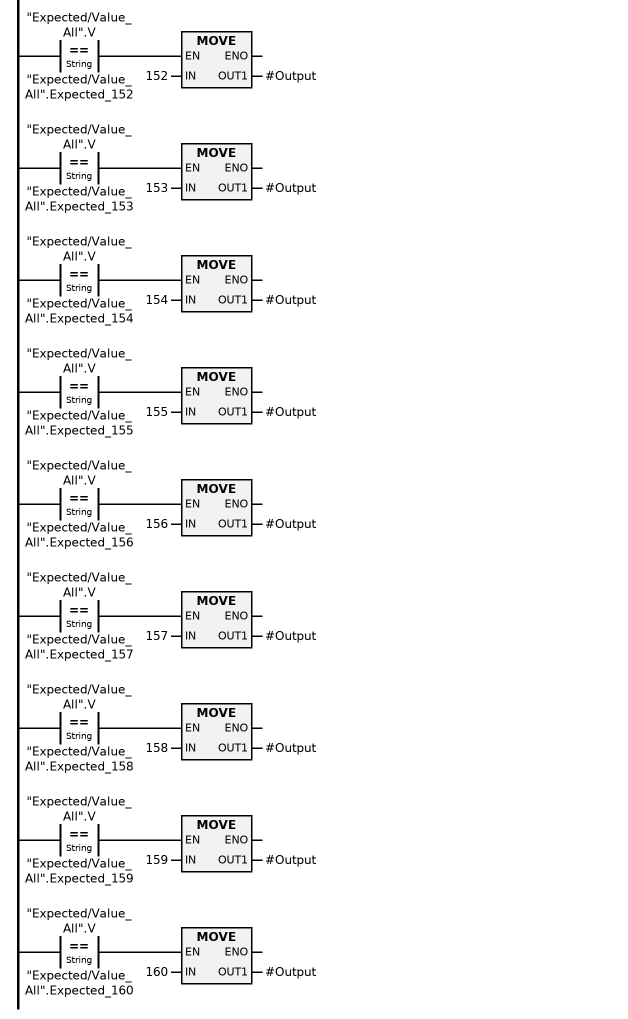
   RUNG wire#powerrail
      { S7_Templates := "SrcType := String" } EQ_Contact(in1 := "Expected/Value_All".V, in2 := "Expected/Value_All".Expected_141)
      Move(in := 141, out1 => #Output)
   END_RUNG
   RUNG wire#powerrail
      { S7_Templates := "SrcType := String" } EQ_Contact(in1 := "Expected/Value_All".V, in2 := "Expected/Value_All".Expected_142)
      Move(in := 142, out1 => #Output)
   END_RUNG
   RUNG wire#powerrail
      { S7_Templates := "SrcType := String" } EQ_Contact(in1 := "Expected/Value_All".V, in2 := "Expected/Value_All".Expected_143)
      Move(in := 143, out1 => #Output)
   END_RUNG
   RUNG wire#powerrail
      { S7_Templates := "SrcType := String" } EQ_Contact(in1 := "Expected/Value_All".V, in2 := "Expected/Value_All".Expected_144)
      Move(in := 144, out1 => #Output)
   END_RUNG
   RUNG wire#powerrail
      { S7_Templates := "SrcType := String" } EQ_Contact(in1 := "Expected/Value_All".V, in2 := "Expected/Value_All".Expected_145)
      Move(in := 145, out1 => #Output)
   END_RUNG
   RUNG wire#powerrail
      { S7_Templates := "SrcType := String" } EQ_Contact(in1 := "Expected/Value_All".V, in2 := "Expected/Value_All".Expected_146)
      Move(in := 146, out1 => #Output)
   END_RUNG
   RUNG wire#powerrail
      { S7_Templates := "SrcType := String" } EQ_Contact(in1 := "Expected/Value_All".V, in2 := "Expected/Value_All".Expected_147)
      Move(in := 147, out1 => #Output)
   END_RUNG
   RUNG wire#powerrail
      { S7_Templates := "SrcType := String" } EQ_Contact(in1 := "Expected/Value_All".V, in2 := "Expected/Value_All".Expected_148)
      Move(in := 148, out1 => #Output)
   END_RUNG
   RUNG wire#powerrail
      { S7_Templates := "SrcType := String" } EQ_Contact(in1 := "Expected/Value_All".V, in2 := "Expected/Value_All".Expected_149)
      Move(in := 149, out1 => #Output)
   END_RUNG
   RUNG wire#powerrail
      { S7_Templates := "SrcType := String" } EQ_Contact(in1 := "Expected/Value_All".V, in2 := "Expected/Value_All".Expected_150)
      Move(in := 150, out1 => #Output)
   END_RUNG
   RUNG wire#powerrail
      { S7_Templates := "SrcType := String" } EQ_Contact(in1 := "Expected/Value_All".V, in2 := "Expected/Value_All".Expected_151)
      Move(in := 151, out1 => #Output)
   END_RUNG
   RUNG wire#powerrail
      { S7_Templates := "SrcType := String" } EQ_Contact(in1 := "Expected/Value_All".V, in2 := "Expected/Value_All".Expected_152)
      Move(in := 152, out1 => #Output)
   END_RUNG
   RUNG wire#powerrail
      { S7_Templates := "SrcType := String" } EQ_Contact(in1 := "Expected/Value_All".V, in2 := "Expected/Value_All".Expected_153)
      Move(in := 153, out1 => #Output)
   END_RUNG
   RUNG wire#powerrail
      { S7_Templates := "SrcType := String" } EQ_Contact(in1 := "Expected/Value_All".V, in2 := "Expected/Value_All".Expected_154)
      Move(in := 154, out1 => #Output)
   END_RUNG
   RUNG wire#powerrail
      { S7_Templates := "SrcType := String" } EQ_Contact(in1 := "Expected/Value_All".V, in2 := "Expected/Value_All".Expected_155)
      Move(in := 155, out1 => #Output)
   END_RUNG
   RUNG wire#powerrail
      { S7_Templates := "SrcType := String" } EQ_Contact(in1 := "Expected/Value_All".V, in2 := "Expected/Value_All".Expected_156)
      Move(in := 156, out1 => #Output)
   END_RUNG
   RUNG wire#powerrail
      { S7_Templates := "SrcType := String" } EQ_Contact(in1 := "Expected/Value_All".V, in2 := "Expected/Value_All".Expected_157)
      Move(in := 157, out1 => #Output)
   END_RUNG
   RUNG wire#powerrail
      { S7_Templates := "SrcType := String" } EQ_Contact(in1 := "Expected/Value_All".V, in2 := "Expected/Value_All".Expected_158)
      Move(in := 158, out1 => #Output)
   END_RUNG
   RUNG wire#powerrail
      { S7_Templates := "SrcType := String" } EQ_Contact(in1 := "Expected/Value_All".V, in2 := "Expected/Value_All".Expected_159)
      Move(in := 159, out1 => #Output)
   END_RUNG
   RUNG wire#powerrail
      { S7_Templates := "SrcType := String" } EQ_Contact(in1 := "Expected/Value_All".V, in2 := "Expected/Value_All".Expected_160)
      Move(in := 160, out1 => #Output)
   END_RUNG
   // the same network as SCL:
   IF "Expected/Value_All".V = "Expected/Value_All".Expected_141 THEN #Output := 141; END_IF;
   IF "Expected/Value_All".V = "Expected/Value_All".Expected_142 THEN #Output := 142; END_IF;
   IF "Expected/Value_All".V = "Expected/Value_All".Expected_143 THEN #Output := 143; END_IF;
   IF "Expected/Value_All".V = "Expected/Value_All".Expected_144 THEN #Output := 144; END_IF;
   IF "Expected/Value_All".V = "Expected/Value_All".Expected_145 THEN #Output := 145; END_IF;
   IF "Expected/Value_All".V = "Expected/Value_All".Expected_146 THEN #Output := 146; END_IF;
   IF "Expected/Value_All".V = "Expected/Value_All".Expected_147 THEN #Output := 147; END_IF;
   IF "Expected/Value_All".V = "Expected/Value_All".Expected_148 THEN #Output := 148; END_IF;
   IF "Expected/Value_All".V = "Expected/Value_All".Expected_149 THEN #Output := 149; END_IF;
   IF "Expected/Value_All".V = "Expected/Value_All".Expected_150 THEN #Output := 150; END_IF;
   IF "Expected/Value_All".V = "Expected/Value_All".Expected_151 THEN #Output := 151; END_IF;
   IF "Expected/Value_All".V = "Expected/Value_All".Expected_152 THEN #Output := 152; END_IF;
   IF "Expected/Value_All".V = "Expected/Value_All".Expected_153 THEN #Output := 153; END_IF;
   IF "Expected/Value_All".V = "Expected/Value_All".Expected_154 THEN #Output := 154; END_IF;
   IF "Expected/Value_All".V = "Expected/Value_All".Expected_155 THEN #Output := 155; END_IF;
   IF "Expected/Value_All".V = "Expected/Value_All".Expected_156 THEN #Output := 156; END_IF;
   IF "Expected/Value_All".V = "Expected/Value_All".Expected_157 THEN #Output := 157; END_IF;
   IF "Expected/Value_All".V = "Expected/Value_All".Expected_158 THEN #Output := 158; END_IF;
   IF "Expected/Value_All".V = "Expected/Value_All".Expected_159 THEN #Output := 159; END_IF;
   IF "Expected/Value_All".V = "Expected/Value_All".Expected_160 THEN #Output := 160; END_IF;
END_REGION

REGION Network 9
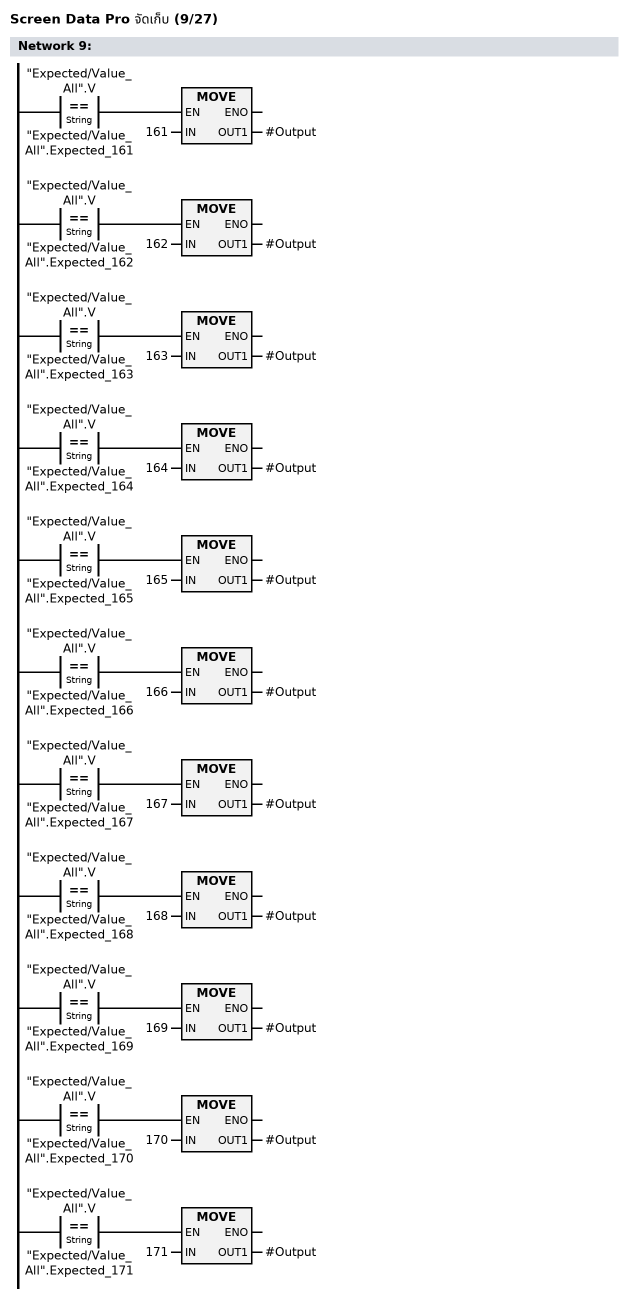
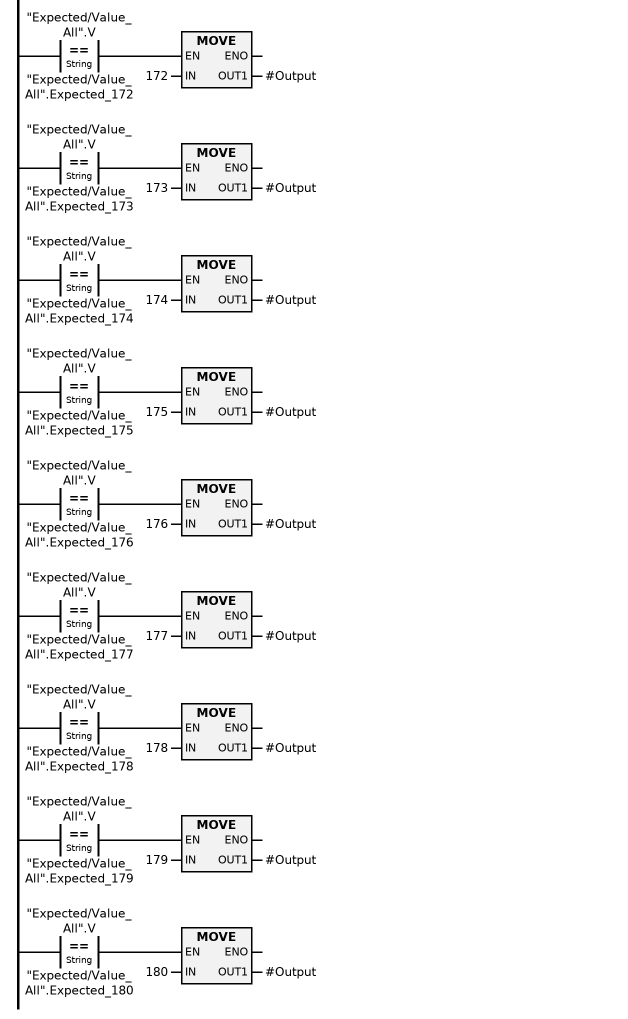
   RUNG wire#powerrail
      { S7_Templates := "SrcType := String" } EQ_Contact(in1 := "Expected/Value_All".V, in2 := "Expected/Value_All".Expected_161)
      Move(in := 161, out1 => #Output)
   END_RUNG
   RUNG wire#powerrail
      { S7_Templates := "SrcType := String" } EQ_Contact(in1 := "Expected/Value_All".V, in2 := "Expected/Value_All".Expected_162)
      Move(in := 162, out1 => #Output)
   END_RUNG
   RUNG wire#powerrail
      { S7_Templates := "SrcType := String" } EQ_Contact(in1 := "Expected/Value_All".V, in2 := "Expected/Value_All".Expected_163)
      Move(in := 163, out1 => #Output)
   END_RUNG
   RUNG wire#powerrail
      { S7_Templates := "SrcType := String" } EQ_Contact(in1 := "Expected/Value_All".V, in2 := "Expected/Value_All".Expected_164)
      Move(in := 164, out1 => #Output)
   END_RUNG
   RUNG wire#powerrail
      { S7_Templates := "SrcType := String" } EQ_Contact(in1 := "Expected/Value_All".V, in2 := "Expected/Value_All".Expected_165)
      Move(in := 165, out1 => #Output)
   END_RUNG
   RUNG wire#powerrail
      { S7_Templates := "SrcType := String" } EQ_Contact(in1 := "Expected/Value_All".V, in2 := "Expected/Value_All".Expected_166)
      Move(in := 166, out1 => #Output)
   END_RUNG
   RUNG wire#powerrail
      { S7_Templates := "SrcType := String" } EQ_Contact(in1 := "Expected/Value_All".V, in2 := "Expected/Value_All".Expected_167)
      Move(in := 167, out1 => #Output)
   END_RUNG
   RUNG wire#powerrail
      { S7_Templates := "SrcType := String" } EQ_Contact(in1 := "Expected/Value_All".V, in2 := "Expected/Value_All".Expected_168)
      Move(in := 168, out1 => #Output)
   END_RUNG
   RUNG wire#powerrail
      { S7_Templates := "SrcType := String" } EQ_Contact(in1 := "Expected/Value_All".V, in2 := "Expected/Value_All".Expected_169)
      Move(in := 169, out1 => #Output)
   END_RUNG
   RUNG wire#powerrail
      { S7_Templates := "SrcType := String" } EQ_Contact(in1 := "Expected/Value_All".V, in2 := "Expected/Value_All".Expected_170)
      Move(in := 170, out1 => #Output)
   END_RUNG
   RUNG wire#powerrail
      { S7_Templates := "SrcType := String" } EQ_Contact(in1 := "Expected/Value_All".V, in2 := "Expected/Value_All".Expected_171)
      Move(in := 171, out1 => #Output)
   END_RUNG
   RUNG wire#powerrail
      { S7_Templates := "SrcType := String" } EQ_Contact(in1 := "Expected/Value_All".V, in2 := "Expected/Value_All".Expected_172)
      Move(in := 172, out1 => #Output)
   END_RUNG
   RUNG wire#powerrail
      { S7_Templates := "SrcType := String" } EQ_Contact(in1 := "Expected/Value_All".V, in2 := "Expected/Value_All".Expected_173)
      Move(in := 173, out1 => #Output)
   END_RUNG
   RUNG wire#powerrail
      { S7_Templates := "SrcType := String" } EQ_Contact(in1 := "Expected/Value_All".V, in2 := "Expected/Value_All".Expected_174)
      Move(in := 174, out1 => #Output)
   END_RUNG
   RUNG wire#powerrail
      { S7_Templates := "SrcType := String" } EQ_Contact(in1 := "Expected/Value_All".V, in2 := "Expected/Value_All".Expected_175)
      Move(in := 175, out1 => #Output)
   END_RUNG
   RUNG wire#powerrail
      { S7_Templates := "SrcType := String" } EQ_Contact(in1 := "Expected/Value_All".V, in2 := "Expected/Value_All".Expected_176)
      Move(in := 176, out1 => #Output)
   END_RUNG
   RUNG wire#powerrail
      { S7_Templates := "SrcType := String" } EQ_Contact(in1 := "Expected/Value_All".V, in2 := "Expected/Value_All".Expected_177)
      Move(in := 177, out1 => #Output)
   END_RUNG
   RUNG wire#powerrail
      { S7_Templates := "SrcType := String" } EQ_Contact(in1 := "Expected/Value_All".V, in2 := "Expected/Value_All".Expected_178)
      Move(in := 178, out1 => #Output)
   END_RUNG
   RUNG wire#powerrail
      { S7_Templates := "SrcType := String" } EQ_Contact(in1 := "Expected/Value_All".V, in2 := "Expected/Value_All".Expected_179)
      Move(in := 179, out1 => #Output)
   END_RUNG
   RUNG wire#powerrail
      { S7_Templates := "SrcType := String" } EQ_Contact(in1 := "Expected/Value_All".V, in2 := "Expected/Value_All".Expected_180)
      Move(in := 180, out1 => #Output)
   END_RUNG
   // the same network as SCL:
   IF "Expected/Value_All".V = "Expected/Value_All".Expected_161 THEN #Output := 161; END_IF;
   IF "Expected/Value_All".V = "Expected/Value_All".Expected_162 THEN #Output := 162; END_IF;
   IF "Expected/Value_All".V = "Expected/Value_All".Expected_163 THEN #Output := 163; END_IF;
   IF "Expected/Value_All".V = "Expected/Value_All".Expected_164 THEN #Output := 164; END_IF;
   IF "Expected/Value_All".V = "Expected/Value_All".Expected_165 THEN #Output := 165; END_IF;
   IF "Expected/Value_All".V = "Expected/Value_All".Expected_166 THEN #Output := 166; END_IF;
   IF "Expected/Value_All".V = "Expected/Value_All".Expected_167 THEN #Output := 167; END_IF;
   IF "Expected/Value_All".V = "Expected/Value_All".Expected_168 THEN #Output := 168; END_IF;
   IF "Expected/Value_All".V = "Expected/Value_All".Expected_169 THEN #Output := 169; END_IF;
   IF "Expected/Value_All".V = "Expected/Value_All".Expected_170 THEN #Output := 170; END_IF;
   IF "Expected/Value_All".V = "Expected/Value_All".Expected_171 THEN #Output := 171; END_IF;
   IF "Expected/Value_All".V = "Expected/Value_All".Expected_172 THEN #Output := 172; END_IF;
   IF "Expected/Value_All".V = "Expected/Value_All".Expected_173 THEN #Output := 173; END_IF;
   IF "Expected/Value_All".V = "Expected/Value_All".Expected_174 THEN #Output := 174; END_IF;
   IF "Expected/Value_All".V = "Expected/Value_All".Expected_175 THEN #Output := 175; END_IF;
   IF "Expected/Value_All".V = "Expected/Value_All".Expected_176 THEN #Output := 176; END_IF;
   IF "Expected/Value_All".V = "Expected/Value_All".Expected_177 THEN #Output := 177; END_IF;
   IF "Expected/Value_All".V = "Expected/Value_All".Expected_178 THEN #Output := 178; END_IF;
   IF "Expected/Value_All".V = "Expected/Value_All".Expected_179 THEN #Output := 179; END_IF;
   IF "Expected/Value_All".V = "Expected/Value_All".Expected_180 THEN #Output := 180; END_IF;
END_REGION

REGION Network 10
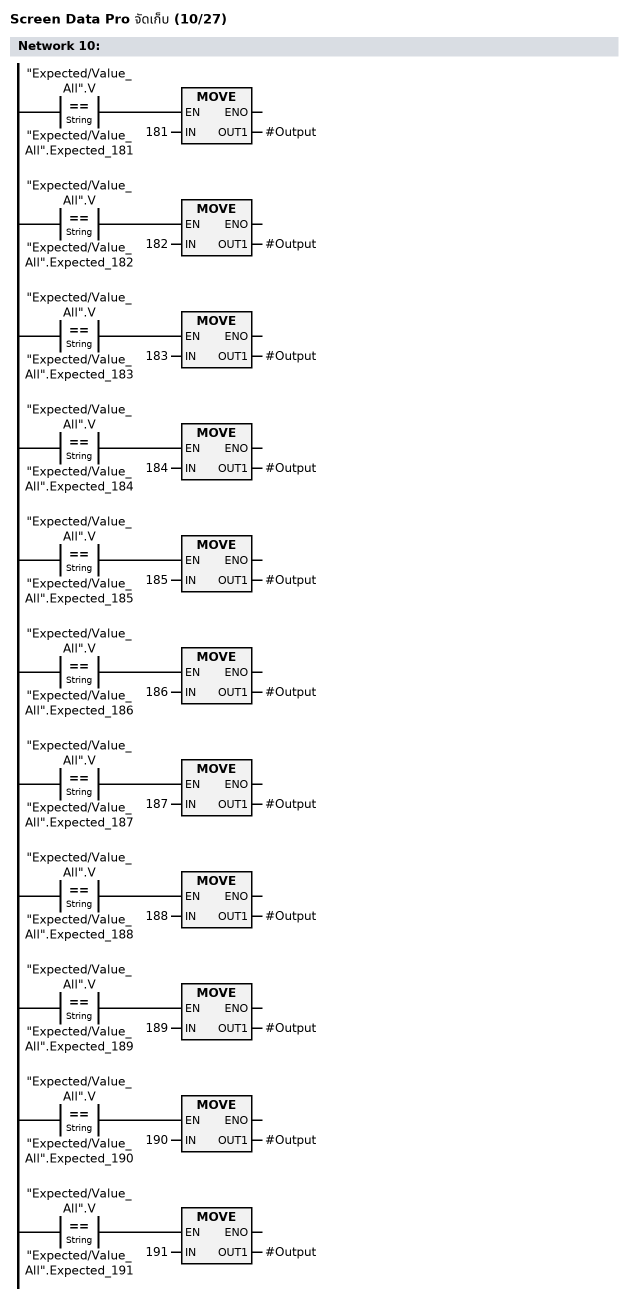
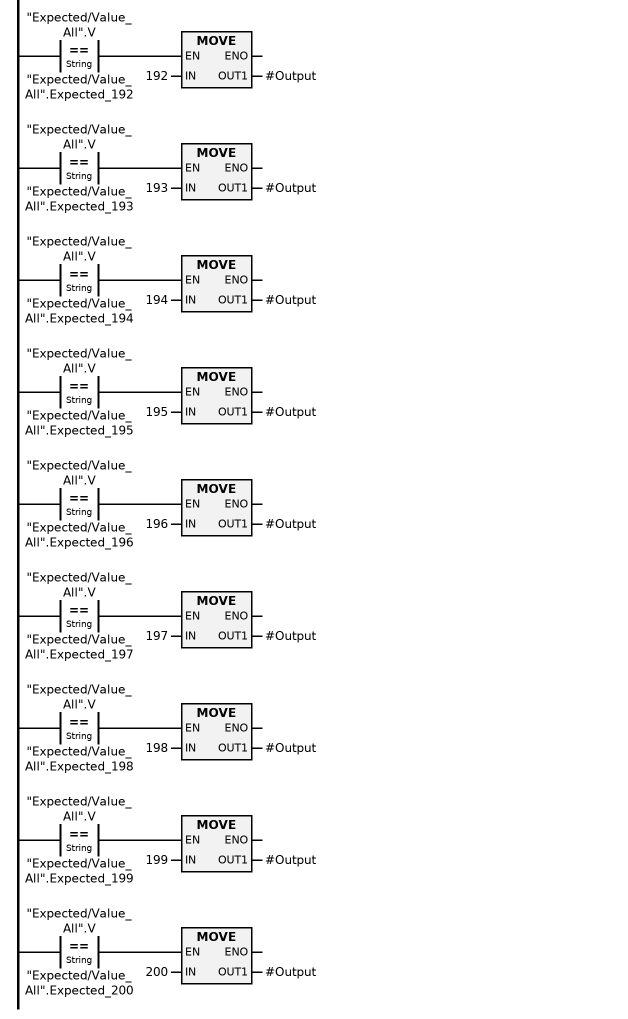
   RUNG wire#powerrail
      { S7_Templates := "SrcType := String" } EQ_Contact(in1 := "Expected/Value_All".V, in2 := "Expected/Value_All".Expected_181)
      Move(in := 181, out1 => #Output)
   END_RUNG
   RUNG wire#powerrail
      { S7_Templates := "SrcType := String" } EQ_Contact(in1 := "Expected/Value_All".V, in2 := "Expected/Value_All".Expected_182)
      Move(in := 182, out1 => #Output)
   END_RUNG
   RUNG wire#powerrail
      { S7_Templates := "SrcType := String" } EQ_Contact(in1 := "Expected/Value_All".V, in2 := "Expected/Value_All".Expected_183)
      Move(in := 183, out1 => #Output)
   END_RUNG
   RUNG wire#powerrail
      { S7_Templates := "SrcType := String" } EQ_Contact(in1 := "Expected/Value_All".V, in2 := "Expected/Value_All".Expected_184)
      Move(in := 184, out1 => #Output)
   END_RUNG
   RUNG wire#powerrail
      { S7_Templates := "SrcType := String" } EQ_Contact(in1 := "Expected/Value_All".V, in2 := "Expected/Value_All".Expected_185)
      Move(in := 185, out1 => #Output)
   END_RUNG
   RUNG wire#powerrail
      { S7_Templates := "SrcType := String" } EQ_Contact(in1 := "Expected/Value_All".V, in2 := "Expected/Value_All".Expected_186)
      Move(in := 186, out1 => #Output)
   END_RUNG
   RUNG wire#powerrail
      { S7_Templates := "SrcType := String" } EQ_Contact(in1 := "Expected/Value_All".V, in2 := "Expected/Value_All".Expected_187)
      Move(in := 187, out1 => #Output)
   END_RUNG
   RUNG wire#powerrail
      { S7_Templates := "SrcType := String" } EQ_Contact(in1 := "Expected/Value_All".V, in2 := "Expected/Value_All".Expected_188)
      Move(in := 188, out1 => #Output)
   END_RUNG
   RUNG wire#powerrail
      { S7_Templates := "SrcType := String" } EQ_Contact(in1 := "Expected/Value_All".V, in2 := "Expected/Value_All".Expected_189)
      Move(in := 189, out1 => #Output)
   END_RUNG
   RUNG wire#powerrail
      { S7_Templates := "SrcType := String" } EQ_Contact(in1 := "Expected/Value_All".V, in2 := "Expected/Value_All".Expected_190)
      Move(in := 190, out1 => #Output)
   END_RUNG
   RUNG wire#powerrail
      { S7_Templates := "SrcType := String" } EQ_Contact(in1 := "Expected/Value_All".V, in2 := "Expected/Value_All".Expected_191)
      Move(in := 191, out1 => #Output)
   END_RUNG
   RUNG wire#powerrail
      { S7_Templates := "SrcType := String" } EQ_Contact(in1 := "Expected/Value_All".V, in2 := "Expected/Value_All".Expected_192)
      Move(in := 192, out1 => #Output)
   END_RUNG
   RUNG wire#powerrail
      { S7_Templates := "SrcType := String" } EQ_Contact(in1 := "Expected/Value_All".V, in2 := "Expected/Value_All".Expected_193)
      Move(in := 193, out1 => #Output)
   END_RUNG
   RUNG wire#powerrail
      { S7_Templates := "SrcType := String" } EQ_Contact(in1 := "Expected/Value_All".V, in2 := "Expected/Value_All".Expected_194)
      Move(in := 194, out1 => #Output)
   END_RUNG
   RUNG wire#powerrail
      { S7_Templates := "SrcType := String" } EQ_Contact(in1 := "Expected/Value_All".V, in2 := "Expected/Value_All".Expected_195)
      Move(in := 195, out1 => #Output)
   END_RUNG
   RUNG wire#powerrail
      { S7_Templates := "SrcType := String" } EQ_Contact(in1 := "Expected/Value_All".V, in2 := "Expected/Value_All".Expected_196)
      Move(in := 196, out1 => #Output)
   END_RUNG
   RUNG wire#powerrail
      { S7_Templates := "SrcType := String" } EQ_Contact(in1 := "Expected/Value_All".V, in2 := "Expected/Value_All".Expected_197)
      Move(in := 197, out1 => #Output)
   END_RUNG
   RUNG wire#powerrail
      { S7_Templates := "SrcType := String" } EQ_Contact(in1 := "Expected/Value_All".V, in2 := "Expected/Value_All".Expected_198)
      Move(in := 198, out1 => #Output)
   END_RUNG
   RUNG wire#powerrail
      { S7_Templates := "SrcType := String" } EQ_Contact(in1 := "Expected/Value_All".V, in2 := "Expected/Value_All".Expected_199)
      Move(in := 199, out1 => #Output)
   END_RUNG
   RUNG wire#powerrail
      { S7_Templates := "SrcType := String" } EQ_Contact(in1 := "Expected/Value_All".V, in2 := "Expected/Value_All".Expected_200)
      Move(in := 200, out1 => #Output)
   END_RUNG
   // the same network as SCL:
   IF "Expected/Value_All".V = "Expected/Value_All".Expected_181 THEN #Output := 181; END_IF;
   IF "Expected/Value_All".V = "Expected/Value_All".Expected_182 THEN #Output := 182; END_IF;
   IF "Expected/Value_All".V = "Expected/Value_All".Expected_183 THEN #Output := 183; END_IF;
   IF "Expected/Value_All".V = "Expected/Value_All".Expected_184 THEN #Output := 184; END_IF;
   IF "Expected/Value_All".V = "Expected/Value_All".Expected_185 THEN #Output := 185; END_IF;
   IF "Expected/Value_All".V = "Expected/Value_All".Expected_186 THEN #Output := 186; END_IF;
   IF "Expected/Value_All".V = "Expected/Value_All".Expected_187 THEN #Output := 187; END_IF;
   IF "Expected/Value_All".V = "Expected/Value_All".Expected_188 THEN #Output := 188; END_IF;
   IF "Expected/Value_All".V = "Expected/Value_All".Expected_189 THEN #Output := 189; END_IF;
   IF "Expected/Value_All".V = "Expected/Value_All".Expected_190 THEN #Output := 190; END_IF;
   IF "Expected/Value_All".V = "Expected/Value_All".Expected_191 THEN #Output := 191; END_IF;
   IF "Expected/Value_All".V = "Expected/Value_All".Expected_192 THEN #Output := 192; END_IF;
   IF "Expected/Value_All".V = "Expected/Value_All".Expected_193 THEN #Output := 193; END_IF;
   IF "Expected/Value_All".V = "Expected/Value_All".Expected_194 THEN #Output := 194; END_IF;
   IF "Expected/Value_All".V = "Expected/Value_All".Expected_195 THEN #Output := 195; END_IF;
   IF "Expected/Value_All".V = "Expected/Value_All".Expected_196 THEN #Output := 196; END_IF;
   IF "Expected/Value_All".V = "Expected/Value_All".Expected_197 THEN #Output := 197; END_IF;
   IF "Expected/Value_All".V = "Expected/Value_All".Expected_198 THEN #Output := 198; END_IF;
   IF "Expected/Value_All".V = "Expected/Value_All".Expected_199 THEN #Output := 199; END_IF;
   IF "Expected/Value_All".V = "Expected/Value_All".Expected_200 THEN #Output := 200; END_IF;
END_REGION

REGION Network 11
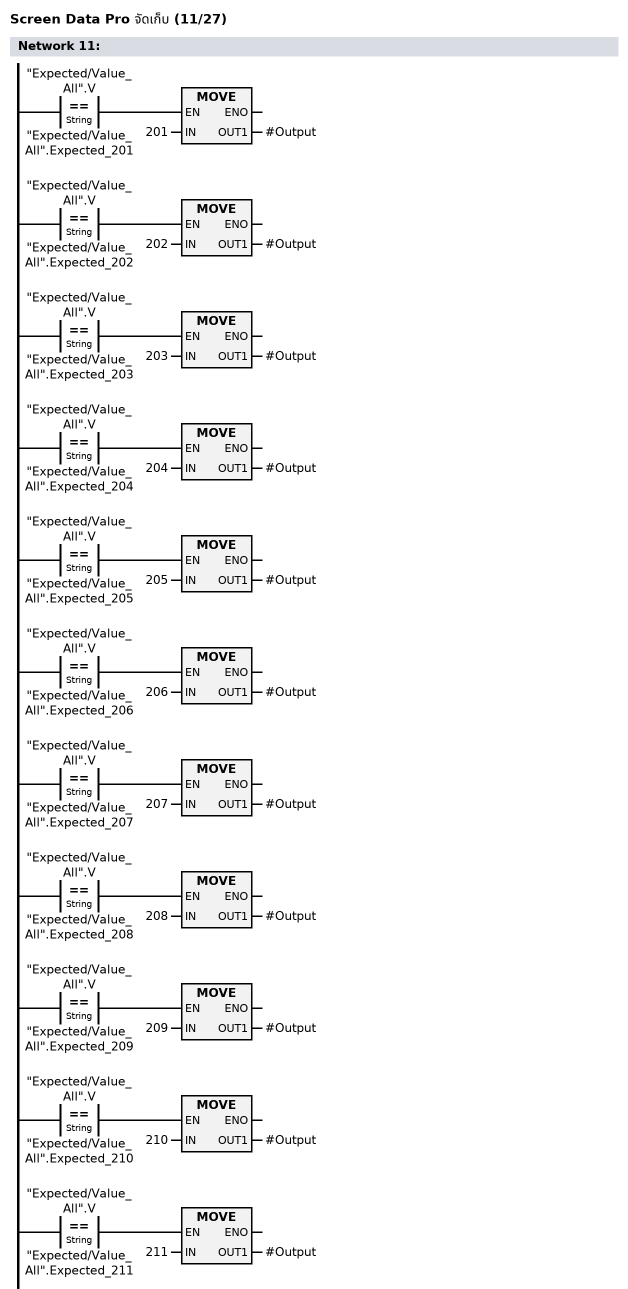
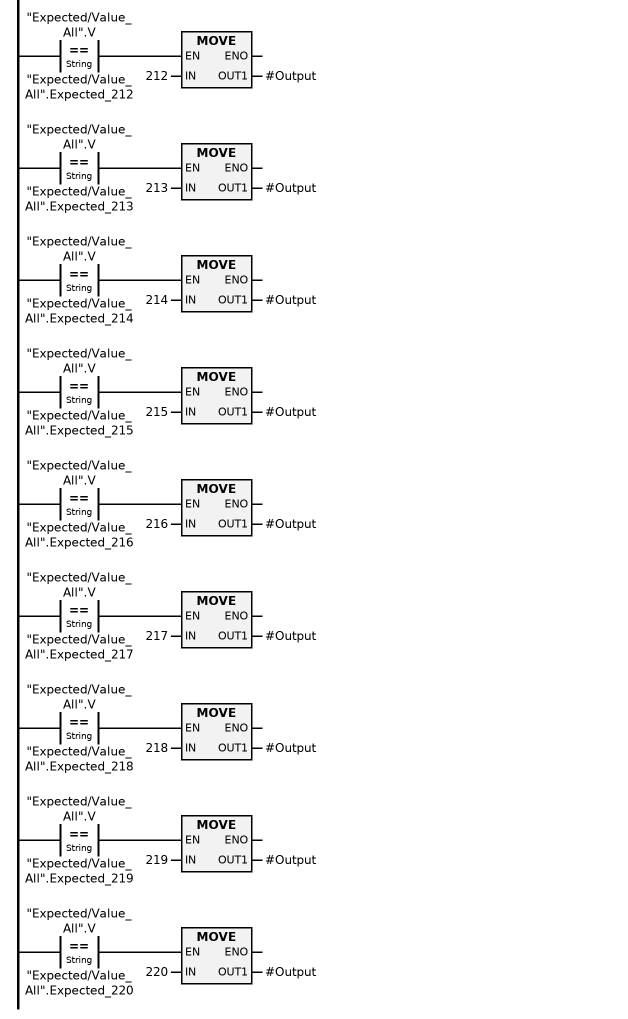
   RUNG wire#powerrail
      { S7_Templates := "SrcType := String" } EQ_Contact(in1 := "Expected/Value_All".V, in2 := "Expected/Value_All".Expected_201)
      Move(in := 201, out1 => #Output)
   END_RUNG
   RUNG wire#powerrail
      { S7_Templates := "SrcType := String" } EQ_Contact(in1 := "Expected/Value_All".V, in2 := "Expected/Value_All".Expected_202)
      Move(in := 202, out1 => #Output)
   END_RUNG
   RUNG wire#powerrail
      { S7_Templates := "SrcType := String" } EQ_Contact(in1 := "Expected/Value_All".V, in2 := "Expected/Value_All".Expected_203)
      Move(in := 203, out1 => #Output)
   END_RUNG
   RUNG wire#powerrail
      { S7_Templates := "SrcType := String" } EQ_Contact(in1 := "Expected/Value_All".V, in2 := "Expected/Value_All".Expected_204)
      Move(in := 204, out1 => #Output)
   END_RUNG
   RUNG wire#powerrail
      { S7_Templates := "SrcType := String" } EQ_Contact(in1 := "Expected/Value_All".V, in2 := "Expected/Value_All".Expected_205)
      Move(in := 205, out1 => #Output)
   END_RUNG
   RUNG wire#powerrail
      { S7_Templates := "SrcType := String" } EQ_Contact(in1 := "Expected/Value_All".V, in2 := "Expected/Value_All".Expected_206)
      Move(in := 206, out1 => #Output)
   END_RUNG
   RUNG wire#powerrail
      { S7_Templates := "SrcType := String" } EQ_Contact(in1 := "Expected/Value_All".V, in2 := "Expected/Value_All".Expected_207)
      Move(in := 207, out1 => #Output)
   END_RUNG
   RUNG wire#powerrail
      { S7_Templates := "SrcType := String" } EQ_Contact(in1 := "Expected/Value_All".V, in2 := "Expected/Value_All".Expected_208)
      Move(in := 208, out1 => #Output)
   END_RUNG
   RUNG wire#powerrail
      { S7_Templates := "SrcType := String" } EQ_Contact(in1 := "Expected/Value_All".V, in2 := "Expected/Value_All".Expected_209)
      Move(in := 209, out1 => #Output)
   END_RUNG
   RUNG wire#powerrail
      { S7_Templates := "SrcType := String" } EQ_Contact(in1 := "Expected/Value_All".V, in2 := "Expected/Value_All".Expected_210)
      Move(in := 210, out1 => #Output)
   END_RUNG
   RUNG wire#powerrail
      { S7_Templates := "SrcType := String" } EQ_Contact(in1 := "Expected/Value_All".V, in2 := "Expected/Value_All".Expected_211)
      Move(in := 211, out1 => #Output)
   END_RUNG
   RUNG wire#powerrail
      { S7_Templates := "SrcType := String" } EQ_Contact(in1 := "Expected/Value_All".V, in2 := "Expected/Value_All".Expected_212)
      Move(in := 212, out1 => #Output)
   END_RUNG
   RUNG wire#powerrail
      { S7_Templates := "SrcType := String" } EQ_Contact(in1 := "Expected/Value_All".V, in2 := "Expected/Value_All".Expected_213)
      Move(in := 213, out1 => #Output)
   END_RUNG
   RUNG wire#powerrail
      { S7_Templates := "SrcType := String" } EQ_Contact(in1 := "Expected/Value_All".V, in2 := "Expected/Value_All".Expected_214)
      Move(in := 214, out1 => #Output)
   END_RUNG
   RUNG wire#powerrail
      { S7_Templates := "SrcType := String" } EQ_Contact(in1 := "Expected/Value_All".V, in2 := "Expected/Value_All".Expected_215)
      Move(in := 215, out1 => #Output)
   END_RUNG
   RUNG wire#powerrail
      { S7_Templates := "SrcType := String" } EQ_Contact(in1 := "Expected/Value_All".V, in2 := "Expected/Value_All".Expected_216)
      Move(in := 216, out1 => #Output)
   END_RUNG
   RUNG wire#powerrail
      { S7_Templates := "SrcType := String" } EQ_Contact(in1 := "Expected/Value_All".V, in2 := "Expected/Value_All".Expected_217)
      Move(in := 217, out1 => #Output)
   END_RUNG
   RUNG wire#powerrail
      { S7_Templates := "SrcType := String" } EQ_Contact(in1 := "Expected/Value_All".V, in2 := "Expected/Value_All".Expected_218)
      Move(in := 218, out1 => #Output)
   END_RUNG
   RUNG wire#powerrail
      { S7_Templates := "SrcType := String" } EQ_Contact(in1 := "Expected/Value_All".V, in2 := "Expected/Value_All".Expected_219)
      Move(in := 219, out1 => #Output)
   END_RUNG
   RUNG wire#powerrail
      { S7_Templates := "SrcType := String" } EQ_Contact(in1 := "Expected/Value_All".V, in2 := "Expected/Value_All".Expected_220)
      Move(in := 220, out1 => #Output)
   END_RUNG
   // the same network as SCL:
   IF "Expected/Value_All".V = "Expected/Value_All".Expected_201 THEN #Output := 201; END_IF;
   IF "Expected/Value_All".V = "Expected/Value_All".Expected_202 THEN #Output := 202; END_IF;
   IF "Expected/Value_All".V = "Expected/Value_All".Expected_203 THEN #Output := 203; END_IF;
   IF "Expected/Value_All".V = "Expected/Value_All".Expected_204 THEN #Output := 204; END_IF;
   IF "Expected/Value_All".V = "Expected/Value_All".Expected_205 THEN #Output := 205; END_IF;
   IF "Expected/Value_All".V = "Expected/Value_All".Expected_206 THEN #Output := 206; END_IF;
   IF "Expected/Value_All".V = "Expected/Value_All".Expected_207 THEN #Output := 207; END_IF;
   IF "Expected/Value_All".V = "Expected/Value_All".Expected_208 THEN #Output := 208; END_IF;
   IF "Expected/Value_All".V = "Expected/Value_All".Expected_209 THEN #Output := 209; END_IF;
   IF "Expected/Value_All".V = "Expected/Value_All".Expected_210 THEN #Output := 210; END_IF;
   IF "Expected/Value_All".V = "Expected/Value_All".Expected_211 THEN #Output := 211; END_IF;
   IF "Expected/Value_All".V = "Expected/Value_All".Expected_212 THEN #Output := 212; END_IF;
   IF "Expected/Value_All".V = "Expected/Value_All".Expected_213 THEN #Output := 213; END_IF;
   IF "Expected/Value_All".V = "Expected/Value_All".Expected_214 THEN #Output := 214; END_IF;
   IF "Expected/Value_All".V = "Expected/Value_All".Expected_215 THEN #Output := 215; END_IF;
   IF "Expected/Value_All".V = "Expected/Value_All".Expected_216 THEN #Output := 216; END_IF;
   IF "Expected/Value_All".V = "Expected/Value_All".Expected_217 THEN #Output := 217; END_IF;
   IF "Expected/Value_All".V = "Expected/Value_All".Expected_218 THEN #Output := 218; END_IF;
   IF "Expected/Value_All".V = "Expected/Value_All".Expected_219 THEN #Output := 219; END_IF;
   IF "Expected/Value_All".V = "Expected/Value_All".Expected_220 THEN #Output := 220; END_IF;
END_REGION

REGION Network 12
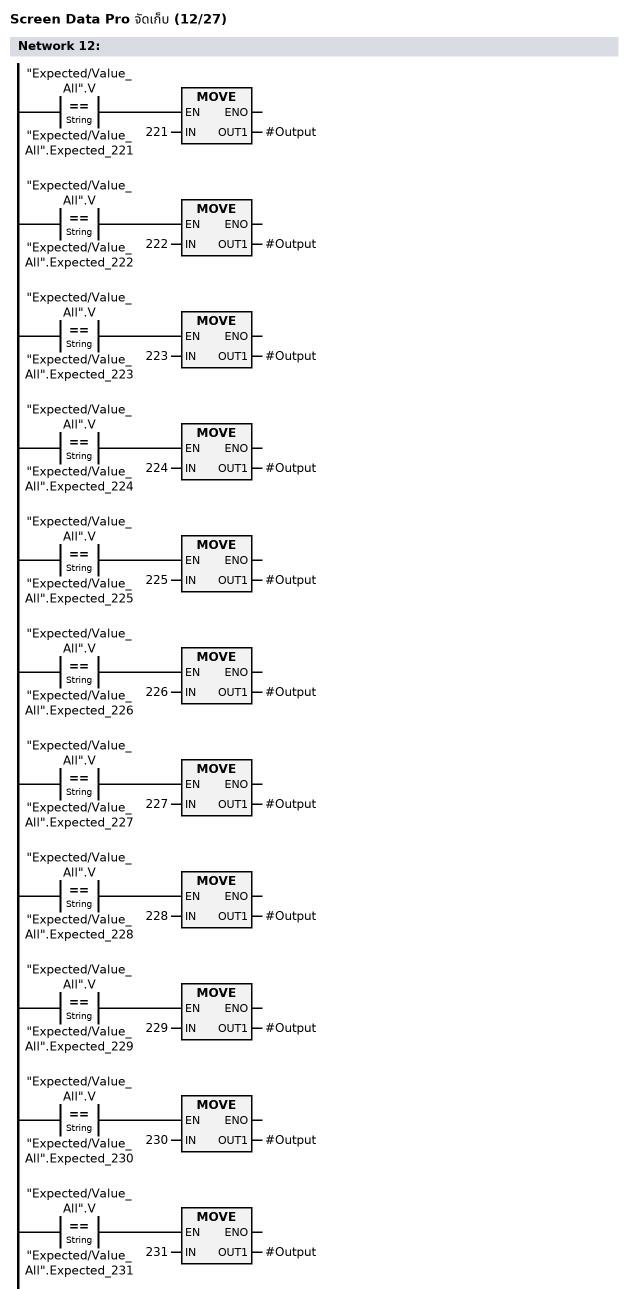
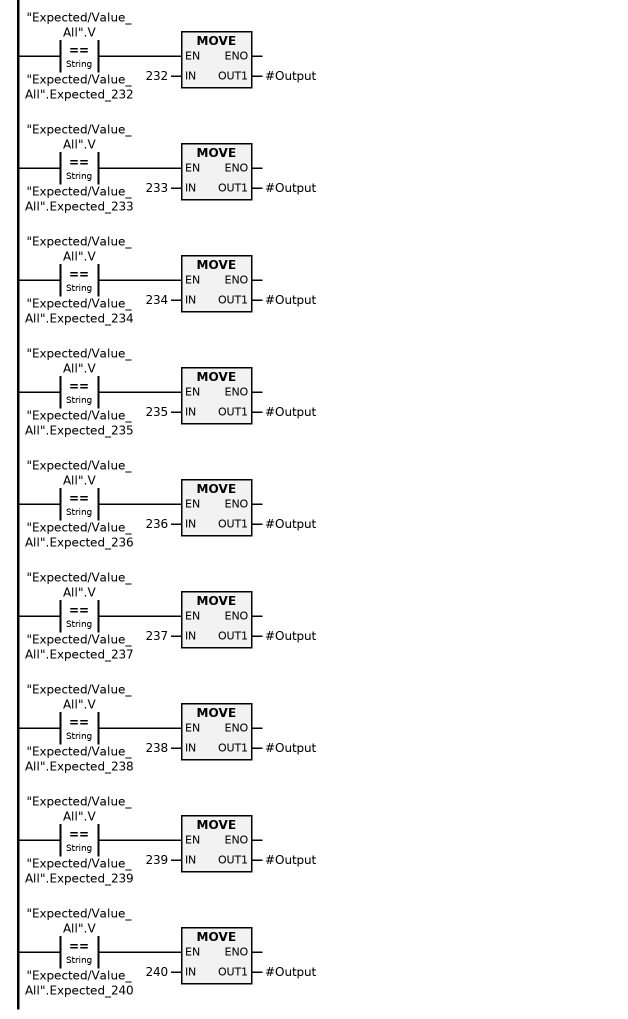
   RUNG wire#powerrail
      { S7_Templates := "SrcType := String" } EQ_Contact(in1 := "Expected/Value_All".V, in2 := "Expected/Value_All".Expected_221)
      Move(in := 221, out1 => #Output)
   END_RUNG
   RUNG wire#powerrail
      { S7_Templates := "SrcType := String" } EQ_Contact(in1 := "Expected/Value_All".V, in2 := "Expected/Value_All".Expected_222)
      Move(in := 222, out1 => #Output)
   END_RUNG
   RUNG wire#powerrail
      { S7_Templates := "SrcType := String" } EQ_Contact(in1 := "Expected/Value_All".V, in2 := "Expected/Value_All".Expected_223)
      Move(in := 223, out1 => #Output)
   END_RUNG
   RUNG wire#powerrail
      { S7_Templates := "SrcType := String" } EQ_Contact(in1 := "Expected/Value_All".V, in2 := "Expected/Value_All".Expected_224)
      Move(in := 224, out1 => #Output)
   END_RUNG
   RUNG wire#powerrail
      { S7_Templates := "SrcType := String" } EQ_Contact(in1 := "Expected/Value_All".V, in2 := "Expected/Value_All".Expected_225)
      Move(in := 225, out1 => #Output)
   END_RUNG
   RUNG wire#powerrail
      { S7_Templates := "SrcType := String" } EQ_Contact(in1 := "Expected/Value_All".V, in2 := "Expected/Value_All".Expected_226)
      Move(in := 226, out1 => #Output)
   END_RUNG
   RUNG wire#powerrail
      { S7_Templates := "SrcType := String" } EQ_Contact(in1 := "Expected/Value_All".V, in2 := "Expected/Value_All".Expected_227)
      Move(in := 227, out1 => #Output)
   END_RUNG
   RUNG wire#powerrail
      { S7_Templates := "SrcType := String" } EQ_Contact(in1 := "Expected/Value_All".V, in2 := "Expected/Value_All".Expected_228)
      Move(in := 228, out1 => #Output)
   END_RUNG
   RUNG wire#powerrail
      { S7_Templates := "SrcType := String" } EQ_Contact(in1 := "Expected/Value_All".V, in2 := "Expected/Value_All".Expected_229)
      Move(in := 229, out1 => #Output)
   END_RUNG
   RUNG wire#powerrail
      { S7_Templates := "SrcType := String" } EQ_Contact(in1 := "Expected/Value_All".V, in2 := "Expected/Value_All".Expected_230)
      Move(in := 230, out1 => #Output)
   END_RUNG
   RUNG wire#powerrail
      { S7_Templates := "SrcType := String" } EQ_Contact(in1 := "Expected/Value_All".V, in2 := "Expected/Value_All".Expected_231)
      Move(in := 231, out1 => #Output)
   END_RUNG
   RUNG wire#powerrail
      { S7_Templates := "SrcType := String" } EQ_Contact(in1 := "Expected/Value_All".V, in2 := "Expected/Value_All".Expected_232)
      Move(in := 232, out1 => #Output)
   END_RUNG
   RUNG wire#powerrail
      { S7_Templates := "SrcType := String" } EQ_Contact(in1 := "Expected/Value_All".V, in2 := "Expected/Value_All".Expected_233)
      Move(in := 233, out1 => #Output)
   END_RUNG
   RUNG wire#powerrail
      { S7_Templates := "SrcType := String" } EQ_Contact(in1 := "Expected/Value_All".V, in2 := "Expected/Value_All".Expected_234)
      Move(in := 234, out1 => #Output)
   END_RUNG
   RUNG wire#powerrail
      { S7_Templates := "SrcType := String" } EQ_Contact(in1 := "Expected/Value_All".V, in2 := "Expected/Value_All".Expected_235)
      Move(in := 235, out1 => #Output)
   END_RUNG
   RUNG wire#powerrail
      { S7_Templates := "SrcType := String" } EQ_Contact(in1 := "Expected/Value_All".V, in2 := "Expected/Value_All".Expected_236)
      Move(in := 236, out1 => #Output)
   END_RUNG
   RUNG wire#powerrail
      { S7_Templates := "SrcType := String" } EQ_Contact(in1 := "Expected/Value_All".V, in2 := "Expected/Value_All".Expected_237)
      Move(in := 237, out1 => #Output)
   END_RUNG
   RUNG wire#powerrail
      { S7_Templates := "SrcType := String" } EQ_Contact(in1 := "Expected/Value_All".V, in2 := "Expected/Value_All".Expected_238)
      Move(in := 238, out1 => #Output)
   END_RUNG
   RUNG wire#powerrail
      { S7_Templates := "SrcType := String" } EQ_Contact(in1 := "Expected/Value_All".V, in2 := "Expected/Value_All".Expected_239)
      Move(in := 239, out1 => #Output)
   END_RUNG
   RUNG wire#powerrail
      { S7_Templates := "SrcType := String" } EQ_Contact(in1 := "Expected/Value_All".V, in2 := "Expected/Value_All".Expected_240)
      Move(in := 240, out1 => #Output)
   END_RUNG
   // the same network as SCL:
   IF "Expected/Value_All".V = "Expected/Value_All".Expected_221 THEN #Output := 221; END_IF;
   IF "Expected/Value_All".V = "Expected/Value_All".Expected_222 THEN #Output := 222; END_IF;
   IF "Expected/Value_All".V = "Expected/Value_All".Expected_223 THEN #Output := 223; END_IF;
   IF "Expected/Value_All".V = "Expected/Value_All".Expected_224 THEN #Output := 224; END_IF;
   IF "Expected/Value_All".V = "Expected/Value_All".Expected_225 THEN #Output := 225; END_IF;
   IF "Expected/Value_All".V = "Expected/Value_All".Expected_226 THEN #Output := 226; END_IF;
   IF "Expected/Value_All".V = "Expected/Value_All".Expected_227 THEN #Output := 227; END_IF;
   IF "Expected/Value_All".V = "Expected/Value_All".Expected_228 THEN #Output := 228; END_IF;
   IF "Expected/Value_All".V = "Expected/Value_All".Expected_229 THEN #Output := 229; END_IF;
   IF "Expected/Value_All".V = "Expected/Value_All".Expected_230 THEN #Output := 230; END_IF;
   IF "Expected/Value_All".V = "Expected/Value_All".Expected_231 THEN #Output := 231; END_IF;
   IF "Expected/Value_All".V = "Expected/Value_All".Expected_232 THEN #Output := 232; END_IF;
   IF "Expected/Value_All".V = "Expected/Value_All".Expected_233 THEN #Output := 233; END_IF;
   IF "Expected/Value_All".V = "Expected/Value_All".Expected_234 THEN #Output := 234; END_IF;
   IF "Expected/Value_All".V = "Expected/Value_All".Expected_235 THEN #Output := 235; END_IF;
   IF "Expected/Value_All".V = "Expected/Value_All".Expected_236 THEN #Output := 236; END_IF;
   IF "Expected/Value_All".V = "Expected/Value_All".Expected_237 THEN #Output := 237; END_IF;
   IF "Expected/Value_All".V = "Expected/Value_All".Expected_238 THEN #Output := 238; END_IF;
   IF "Expected/Value_All".V = "Expected/Value_All".Expected_239 THEN #Output := 239; END_IF;
   IF "Expected/Value_All".V = "Expected/Value_All".Expected_240 THEN #Output := 240; END_IF;
END_REGION

REGION Network 13
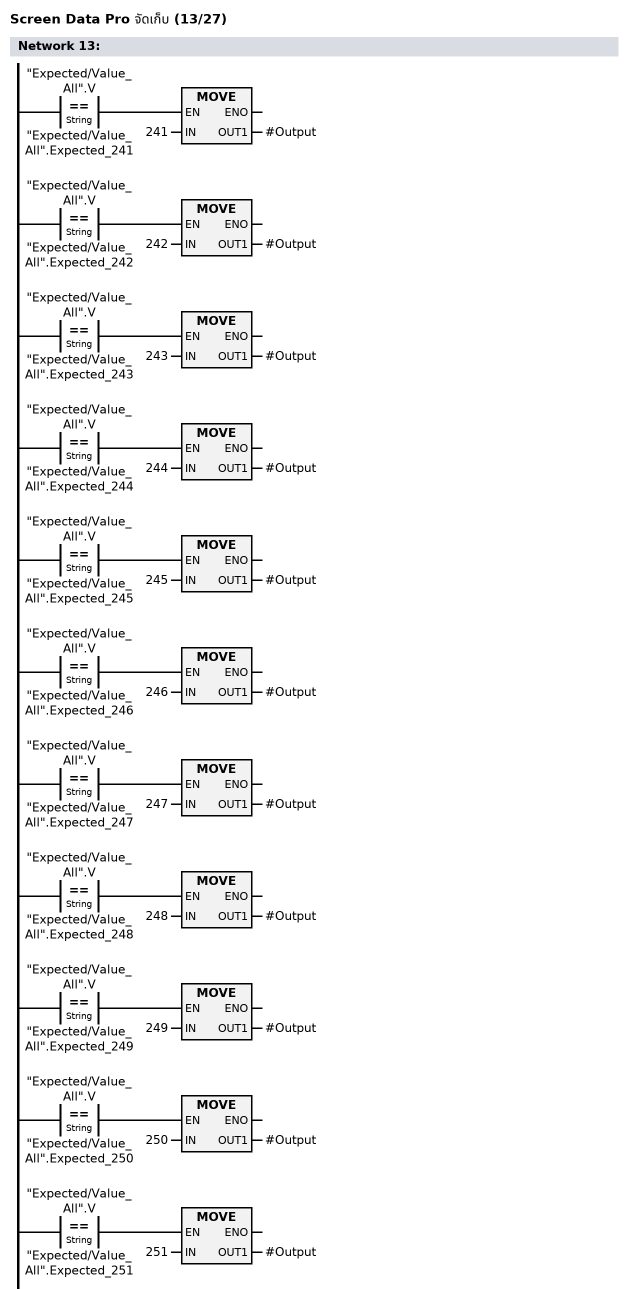
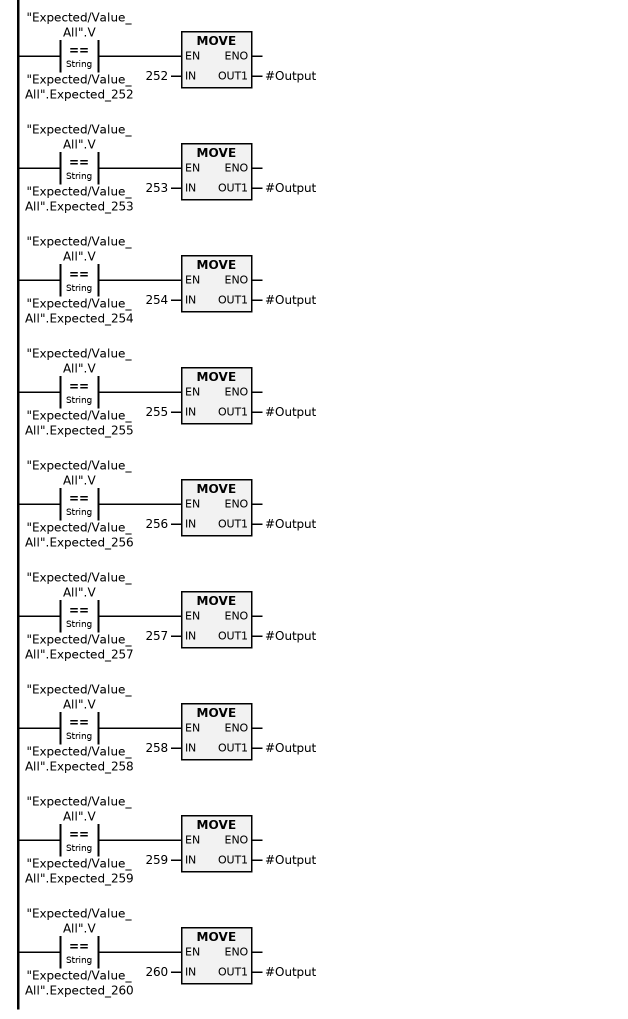
   RUNG wire#powerrail
      { S7_Templates := "SrcType := String" } EQ_Contact(in1 := "Expected/Value_All".V, in2 := "Expected/Value_All".Expected_241)
      Move(in := 241, out1 => #Output)
   END_RUNG
   RUNG wire#powerrail
      { S7_Templates := "SrcType := String" } EQ_Contact(in1 := "Expected/Value_All".V, in2 := "Expected/Value_All".Expected_242)
      Move(in := 242, out1 => #Output)
   END_RUNG
   RUNG wire#powerrail
      { S7_Templates := "SrcType := String" } EQ_Contact(in1 := "Expected/Value_All".V, in2 := "Expected/Value_All".Expected_243)
      Move(in := 243, out1 => #Output)
   END_RUNG
   RUNG wire#powerrail
      { S7_Templates := "SrcType := String" } EQ_Contact(in1 := "Expected/Value_All".V, in2 := "Expected/Value_All".Expected_244)
      Move(in := 244, out1 => #Output)
   END_RUNG
   RUNG wire#powerrail
      { S7_Templates := "SrcType := String" } EQ_Contact(in1 := "Expected/Value_All".V, in2 := "Expected/Value_All".Expected_245)
      Move(in := 245, out1 => #Output)
   END_RUNG
   RUNG wire#powerrail
      { S7_Templates := "SrcType := String" } EQ_Contact(in1 := "Expected/Value_All".V, in2 := "Expected/Value_All".Expected_246)
      Move(in := 246, out1 => #Output)
   END_RUNG
   RUNG wire#powerrail
      { S7_Templates := "SrcType := String" } EQ_Contact(in1 := "Expected/Value_All".V, in2 := "Expected/Value_All".Expected_247)
      Move(in := 247, out1 => #Output)
   END_RUNG
   RUNG wire#powerrail
      { S7_Templates := "SrcType := String" } EQ_Contact(in1 := "Expected/Value_All".V, in2 := "Expected/Value_All".Expected_248)
      Move(in := 248, out1 => #Output)
   END_RUNG
   RUNG wire#powerrail
      { S7_Templates := "SrcType := String" } EQ_Contact(in1 := "Expected/Value_All".V, in2 := "Expected/Value_All".Expected_249)
      Move(in := 249, out1 => #Output)
   END_RUNG
   RUNG wire#powerrail
      { S7_Templates := "SrcType := String" } EQ_Contact(in1 := "Expected/Value_All".V, in2 := "Expected/Value_All".Expected_250)
      Move(in := 250, out1 => #Output)
   END_RUNG
   RUNG wire#powerrail
      { S7_Templates := "SrcType := String" } EQ_Contact(in1 := "Expected/Value_All".V, in2 := "Expected/Value_All".Expected_251)
      Move(in := 251, out1 => #Output)
   END_RUNG
   RUNG wire#powerrail
      { S7_Templates := "SrcType := String" } EQ_Contact(in1 := "Expected/Value_All".V, in2 := "Expected/Value_All".Expected_252)
      Move(in := 252, out1 => #Output)
   END_RUNG
   RUNG wire#powerrail
      { S7_Templates := "SrcType := String" } EQ_Contact(in1 := "Expected/Value_All".V, in2 := "Expected/Value_All".Expected_253)
      Move(in := 253, out1 => #Output)
   END_RUNG
   RUNG wire#powerrail
      { S7_Templates := "SrcType := String" } EQ_Contact(in1 := "Expected/Value_All".V, in2 := "Expected/Value_All".Expected_254)
      Move(in := 254, out1 => #Output)
   END_RUNG
   RUNG wire#powerrail
      { S7_Templates := "SrcType := String" } EQ_Contact(in1 := "Expected/Value_All".V, in2 := "Expected/Value_All".Expected_255)
      Move(in := 255, out1 => #Output)
   END_RUNG
   RUNG wire#powerrail
      { S7_Templates := "SrcType := String" } EQ_Contact(in1 := "Expected/Value_All".V, in2 := "Expected/Value_All".Expected_256)
      Move(in := 256, out1 => #Output)
   END_RUNG
   RUNG wire#powerrail
      { S7_Templates := "SrcType := String" } EQ_Contact(in1 := "Expected/Value_All".V, in2 := "Expected/Value_All".Expected_257)
      Move(in := 257, out1 => #Output)
   END_RUNG
   RUNG wire#powerrail
      { S7_Templates := "SrcType := String" } EQ_Contact(in1 := "Expected/Value_All".V, in2 := "Expected/Value_All".Expected_258)
      Move(in := 258, out1 => #Output)
   END_RUNG
   RUNG wire#powerrail
      { S7_Templates := "SrcType := String" } EQ_Contact(in1 := "Expected/Value_All".V, in2 := "Expected/Value_All".Expected_259)
      Move(in := 259, out1 => #Output)
   END_RUNG
   RUNG wire#powerrail
      { S7_Templates := "SrcType := String" } EQ_Contact(in1 := "Expected/Value_All".V, in2 := "Expected/Value_All".Expected_260)
      Move(in := 260, out1 => #Output)
   END_RUNG
   // the same network as SCL:
   IF "Expected/Value_All".V = "Expected/Value_All".Expected_241 THEN #Output := 241; END_IF;
   IF "Expected/Value_All".V = "Expected/Value_All".Expected_242 THEN #Output := 242; END_IF;
   IF "Expected/Value_All".V = "Expected/Value_All".Expected_243 THEN #Output := 243; END_IF;
   IF "Expected/Value_All".V = "Expected/Value_All".Expected_244 THEN #Output := 244; END_IF;
   IF "Expected/Value_All".V = "Expected/Value_All".Expected_245 THEN #Output := 245; END_IF;
   IF "Expected/Value_All".V = "Expected/Value_All".Expected_246 THEN #Output := 246; END_IF;
   IF "Expected/Value_All".V = "Expected/Value_All".Expected_247 THEN #Output := 247; END_IF;
   IF "Expected/Value_All".V = "Expected/Value_All".Expected_248 THEN #Output := 248; END_IF;
   IF "Expected/Value_All".V = "Expected/Value_All".Expected_249 THEN #Output := 249; END_IF;
   IF "Expected/Value_All".V = "Expected/Value_All".Expected_250 THEN #Output := 250; END_IF;
   IF "Expected/Value_All".V = "Expected/Value_All".Expected_251 THEN #Output := 251; END_IF;
   IF "Expected/Value_All".V = "Expected/Value_All".Expected_252 THEN #Output := 252; END_IF;
   IF "Expected/Value_All".V = "Expected/Value_All".Expected_253 THEN #Output := 253; END_IF;
   IF "Expected/Value_All".V = "Expected/Value_All".Expected_254 THEN #Output := 254; END_IF;
   IF "Expected/Value_All".V = "Expected/Value_All".Expected_255 THEN #Output := 255; END_IF;
   IF "Expected/Value_All".V = "Expected/Value_All".Expected_256 THEN #Output := 256; END_IF;
   IF "Expected/Value_All".V = "Expected/Value_All".Expected_257 THEN #Output := 257; END_IF;
   IF "Expected/Value_All".V = "Expected/Value_All".Expected_258 THEN #Output := 258; END_IF;
   IF "Expected/Value_All".V = "Expected/Value_All".Expected_259 THEN #Output := 259; END_IF;
   IF "Expected/Value_All".V = "Expected/Value_All".Expected_260 THEN #Output := 260; END_IF;
END_REGION

REGION Network 14
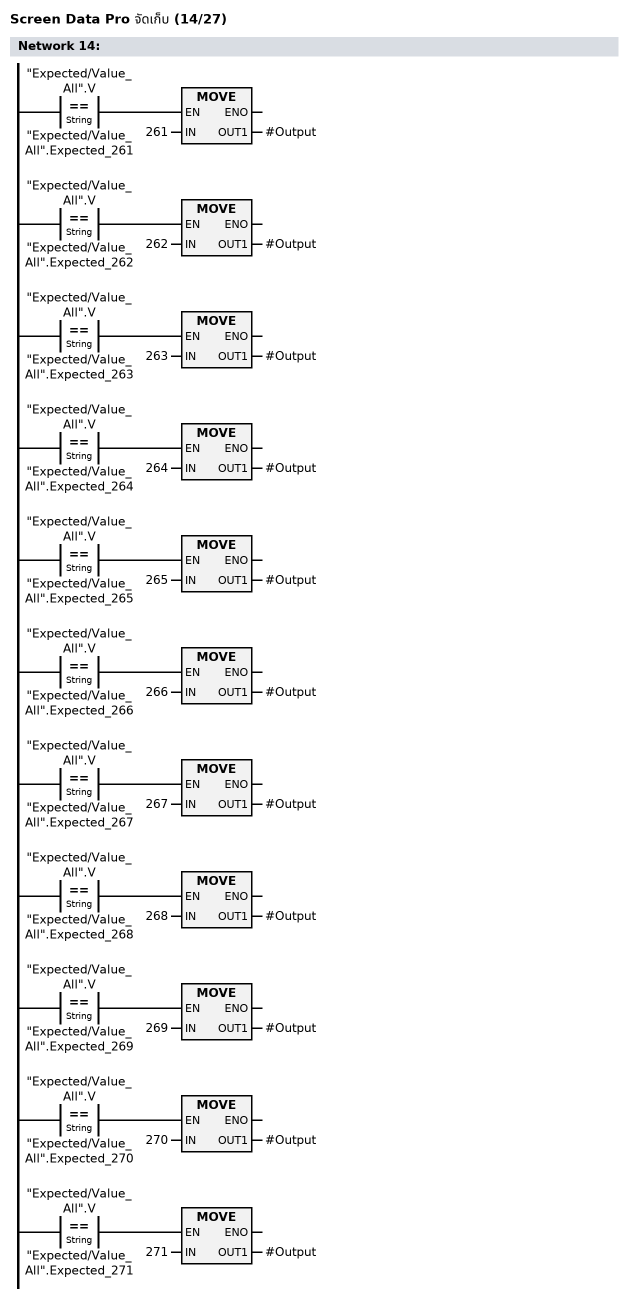
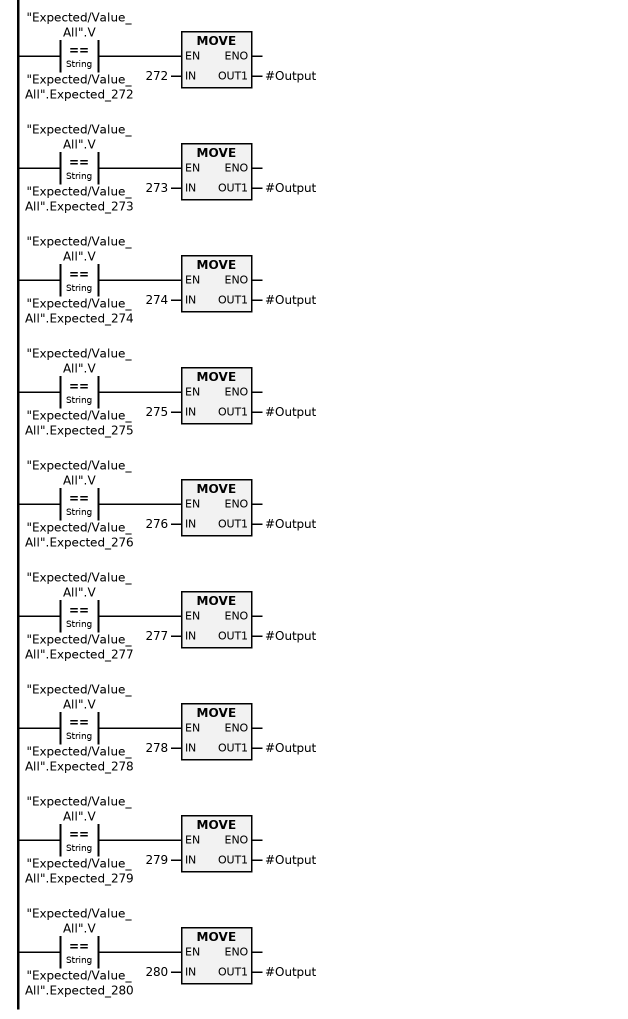
   RUNG wire#powerrail
      { S7_Templates := "SrcType := String" } EQ_Contact(in1 := "Expected/Value_All".V, in2 := "Expected/Value_All".Expected_261)
      Move(in := 261, out1 => #Output)
   END_RUNG
   RUNG wire#powerrail
      { S7_Templates := "SrcType := String" } EQ_Contact(in1 := "Expected/Value_All".V, in2 := "Expected/Value_All".Expected_262)
      Move(in := 262, out1 => #Output)
   END_RUNG
   RUNG wire#powerrail
      { S7_Templates := "SrcType := String" } EQ_Contact(in1 := "Expected/Value_All".V, in2 := "Expected/Value_All".Expected_263)
      Move(in := 263, out1 => #Output)
   END_RUNG
   RUNG wire#powerrail
      { S7_Templates := "SrcType := String" } EQ_Contact(in1 := "Expected/Value_All".V, in2 := "Expected/Value_All".Expected_264)
      Move(in := 264, out1 => #Output)
   END_RUNG
   RUNG wire#powerrail
      { S7_Templates := "SrcType := String" } EQ_Contact(in1 := "Expected/Value_All".V, in2 := "Expected/Value_All".Expected_265)
      Move(in := 265, out1 => #Output)
   END_RUNG
   RUNG wire#powerrail
      { S7_Templates := "SrcType := String" } EQ_Contact(in1 := "Expected/Value_All".V, in2 := "Expected/Value_All".Expected_266)
      Move(in := 266, out1 => #Output)
   END_RUNG
   RUNG wire#powerrail
      { S7_Templates := "SrcType := String" } EQ_Contact(in1 := "Expected/Value_All".V, in2 := "Expected/Value_All".Expected_267)
      Move(in := 267, out1 => #Output)
   END_RUNG
   RUNG wire#powerrail
      { S7_Templates := "SrcType := String" } EQ_Contact(in1 := "Expected/Value_All".V, in2 := "Expected/Value_All".Expected_268)
      Move(in := 268, out1 => #Output)
   END_RUNG
   RUNG wire#powerrail
      { S7_Templates := "SrcType := String" } EQ_Contact(in1 := "Expected/Value_All".V, in2 := "Expected/Value_All".Expected_269)
      Move(in := 269, out1 => #Output)
   END_RUNG
   RUNG wire#powerrail
      { S7_Templates := "SrcType := String" } EQ_Contact(in1 := "Expected/Value_All".V, in2 := "Expected/Value_All".Expected_270)
      Move(in := 270, out1 => #Output)
   END_RUNG
   RUNG wire#powerrail
      { S7_Templates := "SrcType := String" } EQ_Contact(in1 := "Expected/Value_All".V, in2 := "Expected/Value_All".Expected_271)
      Move(in := 271, out1 => #Output)
   END_RUNG
   RUNG wire#powerrail
      { S7_Templates := "SrcType := String" } EQ_Contact(in1 := "Expected/Value_All".V, in2 := "Expected/Value_All".Expected_272)
      Move(in := 272, out1 => #Output)
   END_RUNG
   RUNG wire#powerrail
      { S7_Templates := "SrcType := String" } EQ_Contact(in1 := "Expected/Value_All".V, in2 := "Expected/Value_All".Expected_273)
      Move(in := 273, out1 => #Output)
   END_RUNG
   RUNG wire#powerrail
      { S7_Templates := "SrcType := String" } EQ_Contact(in1 := "Expected/Value_All".V, in2 := "Expected/Value_All".Expected_274)
      Move(in := 274, out1 => #Output)
   END_RUNG
   RUNG wire#powerrail
      { S7_Templates := "SrcType := String" } EQ_Contact(in1 := "Expected/Value_All".V, in2 := "Expected/Value_All".Expected_275)
      Move(in := 275, out1 => #Output)
   END_RUNG
   RUNG wire#powerrail
      { S7_Templates := "SrcType := String" } EQ_Contact(in1 := "Expected/Value_All".V, in2 := "Expected/Value_All".Expected_276)
      Move(in := 276, out1 => #Output)
   END_RUNG
   RUNG wire#powerrail
      { S7_Templates := "SrcType := String" } EQ_Contact(in1 := "Expected/Value_All".V, in2 := "Expected/Value_All".Expected_277)
      Move(in := 277, out1 => #Output)
   END_RUNG
   RUNG wire#powerrail
      { S7_Templates := "SrcType := String" } EQ_Contact(in1 := "Expected/Value_All".V, in2 := "Expected/Value_All".Expected_278)
      Move(in := 278, out1 => #Output)
   END_RUNG
   RUNG wire#powerrail
      { S7_Templates := "SrcType := String" } EQ_Contact(in1 := "Expected/Value_All".V, in2 := "Expected/Value_All".Expected_279)
      Move(in := 279, out1 => #Output)
   END_RUNG
   RUNG wire#powerrail
      { S7_Templates := "SrcType := String" } EQ_Contact(in1 := "Expected/Value_All".V, in2 := "Expected/Value_All".Expected_280)
      Move(in := 280, out1 => #Output)
   END_RUNG
   // the same network as SCL:
   IF "Expected/Value_All".V = "Expected/Value_All".Expected_261 THEN #Output := 261; END_IF;
   IF "Expected/Value_All".V = "Expected/Value_All".Expected_262 THEN #Output := 262; END_IF;
   IF "Expected/Value_All".V = "Expected/Value_All".Expected_263 THEN #Output := 263; END_IF;
   IF "Expected/Value_All".V = "Expected/Value_All".Expected_264 THEN #Output := 264; END_IF;
   IF "Expected/Value_All".V = "Expected/Value_All".Expected_265 THEN #Output := 265; END_IF;
   IF "Expected/Value_All".V = "Expected/Value_All".Expected_266 THEN #Output := 266; END_IF;
   IF "Expected/Value_All".V = "Expected/Value_All".Expected_267 THEN #Output := 267; END_IF;
   IF "Expected/Value_All".V = "Expected/Value_All".Expected_268 THEN #Output := 268; END_IF;
   IF "Expected/Value_All".V = "Expected/Value_All".Expected_269 THEN #Output := 269; END_IF;
   IF "Expected/Value_All".V = "Expected/Value_All".Expected_270 THEN #Output := 270; END_IF;
   IF "Expected/Value_All".V = "Expected/Value_All".Expected_271 THEN #Output := 271; END_IF;
   IF "Expected/Value_All".V = "Expected/Value_All".Expected_272 THEN #Output := 272; END_IF;
   IF "Expected/Value_All".V = "Expected/Value_All".Expected_273 THEN #Output := 273; END_IF;
   IF "Expected/Value_All".V = "Expected/Value_All".Expected_274 THEN #Output := 274; END_IF;
   IF "Expected/Value_All".V = "Expected/Value_All".Expected_275 THEN #Output := 275; END_IF;
   IF "Expected/Value_All".V = "Expected/Value_All".Expected_276 THEN #Output := 276; END_IF;
   IF "Expected/Value_All".V = "Expected/Value_All".Expected_277 THEN #Output := 277; END_IF;
   IF "Expected/Value_All".V = "Expected/Value_All".Expected_278 THEN #Output := 278; END_IF;
   IF "Expected/Value_All".V = "Expected/Value_All".Expected_279 THEN #Output := 279; END_IF;
   IF "Expected/Value_All".V = "Expected/Value_All".Expected_280 THEN #Output := 280; END_IF;
END_REGION

REGION Network 15
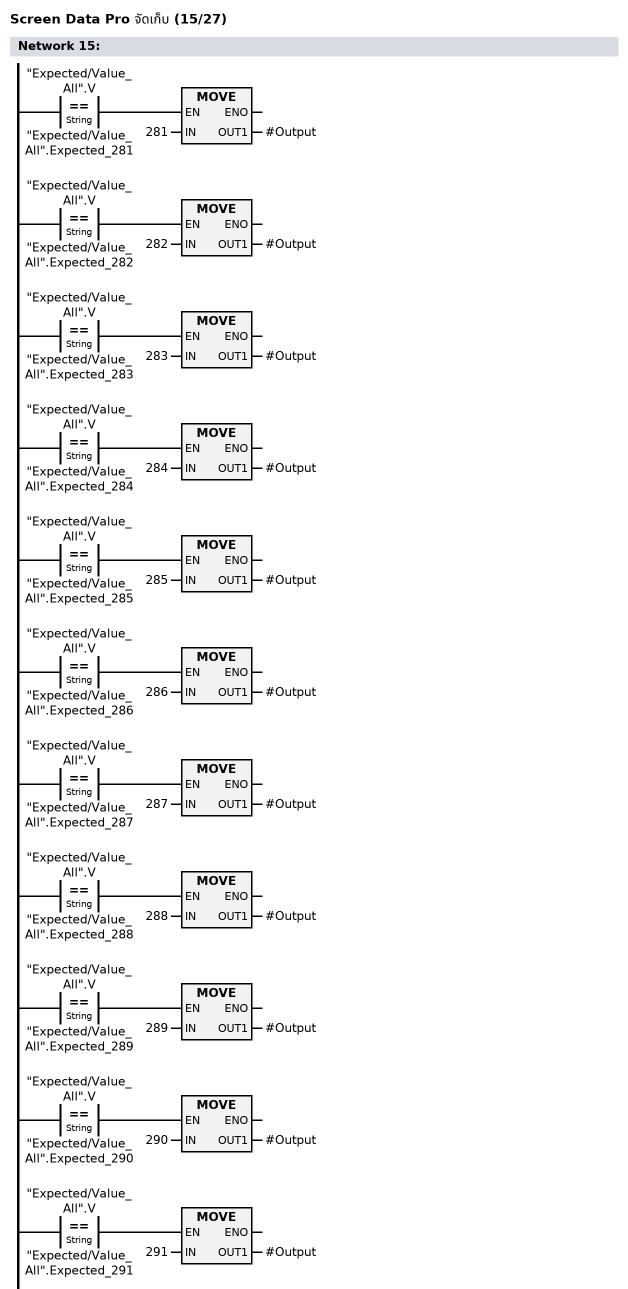
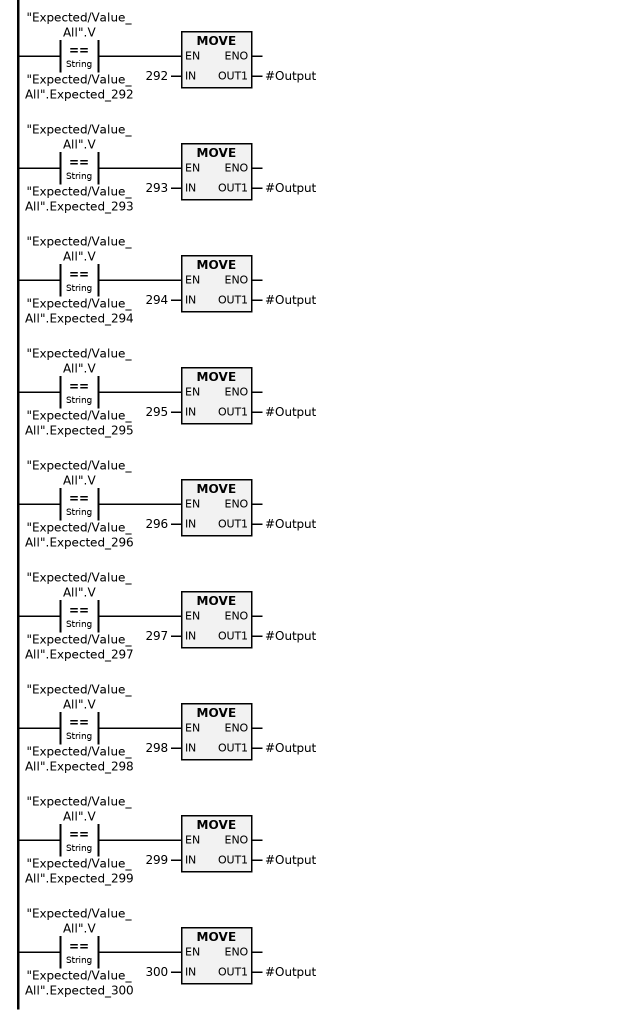
   RUNG wire#powerrail
      { S7_Templates := "SrcType := String" } EQ_Contact(in1 := "Expected/Value_All".V, in2 := "Expected/Value_All".Expected_281)
      Move(in := 281, out1 => #Output)
   END_RUNG
   RUNG wire#powerrail
      { S7_Templates := "SrcType := String" } EQ_Contact(in1 := "Expected/Value_All".V, in2 := "Expected/Value_All".Expected_282)
      Move(in := 282, out1 => #Output)
   END_RUNG
   RUNG wire#powerrail
      { S7_Templates := "SrcType := String" } EQ_Contact(in1 := "Expected/Value_All".V, in2 := "Expected/Value_All".Expected_283)
      Move(in := 283, out1 => #Output)
   END_RUNG
   RUNG wire#powerrail
      { S7_Templates := "SrcType := String" } EQ_Contact(in1 := "Expected/Value_All".V, in2 := "Expected/Value_All".Expected_284)
      Move(in := 284, out1 => #Output)
   END_RUNG
   RUNG wire#powerrail
      { S7_Templates := "SrcType := String" } EQ_Contact(in1 := "Expected/Value_All".V, in2 := "Expected/Value_All".Expected_285)
      Move(in := 285, out1 => #Output)
   END_RUNG
   RUNG wire#powerrail
      { S7_Templates := "SrcType := String" } EQ_Contact(in1 := "Expected/Value_All".V, in2 := "Expected/Value_All".Expected_286)
      Move(in := 286, out1 => #Output)
   END_RUNG
   RUNG wire#powerrail
      { S7_Templates := "SrcType := String" } EQ_Contact(in1 := "Expected/Value_All".V, in2 := "Expected/Value_All".Expected_287)
      Move(in := 287, out1 => #Output)
   END_RUNG
   RUNG wire#powerrail
      { S7_Templates := "SrcType := String" } EQ_Contact(in1 := "Expected/Value_All".V, in2 := "Expected/Value_All".Expected_288)
      Move(in := 288, out1 => #Output)
   END_RUNG
   RUNG wire#powerrail
      { S7_Templates := "SrcType := String" } EQ_Contact(in1 := "Expected/Value_All".V, in2 := "Expected/Value_All".Expected_289)
      Move(in := 289, out1 => #Output)
   END_RUNG
   RUNG wire#powerrail
      { S7_Templates := "SrcType := String" } EQ_Contact(in1 := "Expected/Value_All".V, in2 := "Expected/Value_All".Expected_290)
      Move(in := 290, out1 => #Output)
   END_RUNG
   RUNG wire#powerrail
      { S7_Templates := "SrcType := String" } EQ_Contact(in1 := "Expected/Value_All".V, in2 := "Expected/Value_All".Expected_291)
      Move(in := 291, out1 => #Output)
   END_RUNG
   RUNG wire#powerrail
      { S7_Templates := "SrcType := String" } EQ_Contact(in1 := "Expected/Value_All".V, in2 := "Expected/Value_All".Expected_292)
      Move(in := 292, out1 => #Output)
   END_RUNG
   RUNG wire#powerrail
      { S7_Templates := "SrcType := String" } EQ_Contact(in1 := "Expected/Value_All".V, in2 := "Expected/Value_All".Expected_293)
      Move(in := 293, out1 => #Output)
   END_RUNG
   RUNG wire#powerrail
      { S7_Templates := "SrcType := String" } EQ_Contact(in1 := "Expected/Value_All".V, in2 := "Expected/Value_All".Expected_294)
      Move(in := 294, out1 => #Output)
   END_RUNG
   RUNG wire#powerrail
      { S7_Templates := "SrcType := String" } EQ_Contact(in1 := "Expected/Value_All".V, in2 := "Expected/Value_All".Expected_295)
      Move(in := 295, out1 => #Output)
   END_RUNG
   RUNG wire#powerrail
      { S7_Templates := "SrcType := String" } EQ_Contact(in1 := "Expected/Value_All".V, in2 := "Expected/Value_All".Expected_296)
      Move(in := 296, out1 => #Output)
   END_RUNG
   RUNG wire#powerrail
      { S7_Templates := "SrcType := String" } EQ_Contact(in1 := "Expected/Value_All".V, in2 := "Expected/Value_All".Expected_297)
      Move(in := 297, out1 => #Output)
   END_RUNG
   RUNG wire#powerrail
      { S7_Templates := "SrcType := String" } EQ_Contact(in1 := "Expected/Value_All".V, in2 := "Expected/Value_All".Expected_298)
      Move(in := 298, out1 => #Output)
   END_RUNG
   RUNG wire#powerrail
      { S7_Templates := "SrcType := String" } EQ_Contact(in1 := "Expected/Value_All".V, in2 := "Expected/Value_All".Expected_299)
      Move(in := 299, out1 => #Output)
   END_RUNG
   RUNG wire#powerrail
      { S7_Templates := "SrcType := String" } EQ_Contact(in1 := "Expected/Value_All".V, in2 := "Expected/Value_All".Expected_300)
      Move(in := 300, out1 => #Output)
   END_RUNG
   // the same network as SCL:
   IF "Expected/Value_All".V = "Expected/Value_All".Expected_281 THEN #Output := 281; END_IF;
   IF "Expected/Value_All".V = "Expected/Value_All".Expected_282 THEN #Output := 282; END_IF;
   IF "Expected/Value_All".V = "Expected/Value_All".Expected_283 THEN #Output := 283; END_IF;
   IF "Expected/Value_All".V = "Expected/Value_All".Expected_284 THEN #Output := 284; END_IF;
   IF "Expected/Value_All".V = "Expected/Value_All".Expected_285 THEN #Output := 285; END_IF;
   IF "Expected/Value_All".V = "Expected/Value_All".Expected_286 THEN #Output := 286; END_IF;
   IF "Expected/Value_All".V = "Expected/Value_All".Expected_287 THEN #Output := 287; END_IF;
   IF "Expected/Value_All".V = "Expected/Value_All".Expected_288 THEN #Output := 288; END_IF;
   IF "Expected/Value_All".V = "Expected/Value_All".Expected_289 THEN #Output := 289; END_IF;
   IF "Expected/Value_All".V = "Expected/Value_All".Expected_290 THEN #Output := 290; END_IF;
   IF "Expected/Value_All".V = "Expected/Value_All".Expected_291 THEN #Output := 291; END_IF;
   IF "Expected/Value_All".V = "Expected/Value_All".Expected_292 THEN #Output := 292; END_IF;
   IF "Expected/Value_All".V = "Expected/Value_All".Expected_293 THEN #Output := 293; END_IF;
   IF "Expected/Value_All".V = "Expected/Value_All".Expected_294 THEN #Output := 294; END_IF;
   IF "Expected/Value_All".V = "Expected/Value_All".Expected_295 THEN #Output := 295; END_IF;
   IF "Expected/Value_All".V = "Expected/Value_All".Expected_296 THEN #Output := 296; END_IF;
   IF "Expected/Value_All".V = "Expected/Value_All".Expected_297 THEN #Output := 297; END_IF;
   IF "Expected/Value_All".V = "Expected/Value_All".Expected_298 THEN #Output := 298; END_IF;
   IF "Expected/Value_All".V = "Expected/Value_All".Expected_299 THEN #Output := 299; END_IF;
   IF "Expected/Value_All".V = "Expected/Value_All".Expected_300 THEN #Output := 300; END_IF;
END_REGION

REGION Network 16
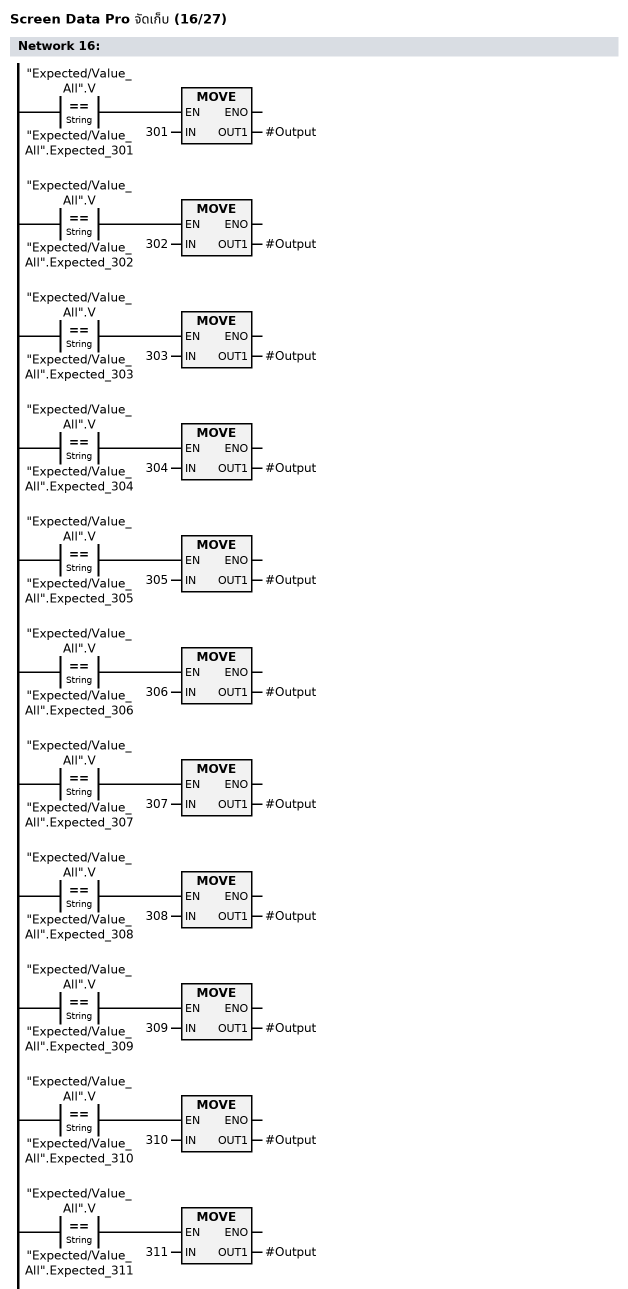
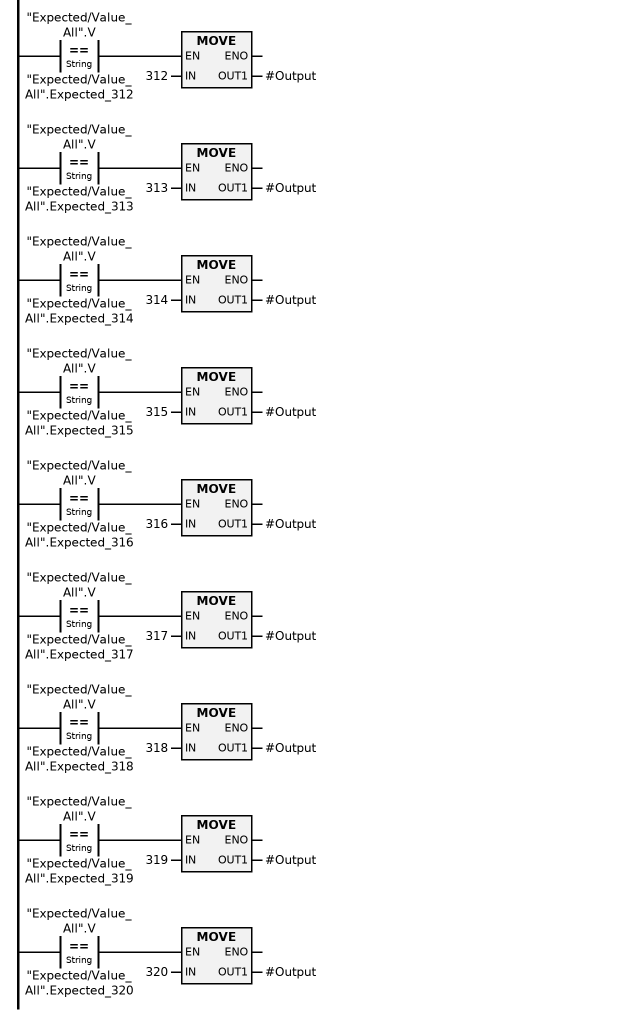
   RUNG wire#powerrail
      { S7_Templates := "SrcType := String" } EQ_Contact(in1 := "Expected/Value_All".V, in2 := "Expected/Value_All".Expected_301)
      Move(in := 301, out1 => #Output)
   END_RUNG
   RUNG wire#powerrail
      { S7_Templates := "SrcType := String" } EQ_Contact(in1 := "Expected/Value_All".V, in2 := "Expected/Value_All".Expected_302)
      Move(in := 302, out1 => #Output)
   END_RUNG
   RUNG wire#powerrail
      { S7_Templates := "SrcType := String" } EQ_Contact(in1 := "Expected/Value_All".V, in2 := "Expected/Value_All".Expected_303)
      Move(in := 303, out1 => #Output)
   END_RUNG
   RUNG wire#powerrail
      { S7_Templates := "SrcType := String" } EQ_Contact(in1 := "Expected/Value_All".V, in2 := "Expected/Value_All".Expected_304)
      Move(in := 304, out1 => #Output)
   END_RUNG
   RUNG wire#powerrail
      { S7_Templates := "SrcType := String" } EQ_Contact(in1 := "Expected/Value_All".V, in2 := "Expected/Value_All".Expected_305)
      Move(in := 305, out1 => #Output)
   END_RUNG
   RUNG wire#powerrail
      { S7_Templates := "SrcType := String" } EQ_Contact(in1 := "Expected/Value_All".V, in2 := "Expected/Value_All".Expected_306)
      Move(in := 306, out1 => #Output)
   END_RUNG
   RUNG wire#powerrail
      { S7_Templates := "SrcType := String" } EQ_Contact(in1 := "Expected/Value_All".V, in2 := "Expected/Value_All".Expected_307)
      Move(in := 307, out1 => #Output)
   END_RUNG
   RUNG wire#powerrail
      { S7_Templates := "SrcType := String" } EQ_Contact(in1 := "Expected/Value_All".V, in2 := "Expected/Value_All".Expected_308)
      Move(in := 308, out1 => #Output)
   END_RUNG
   RUNG wire#powerrail
      { S7_Templates := "SrcType := String" } EQ_Contact(in1 := "Expected/Value_All".V, in2 := "Expected/Value_All".Expected_309)
      Move(in := 309, out1 => #Output)
   END_RUNG
   RUNG wire#powerrail
      { S7_Templates := "SrcType := String" } EQ_Contact(in1 := "Expected/Value_All".V, in2 := "Expected/Value_All".Expected_310)
      Move(in := 310, out1 => #Output)
   END_RUNG
   RUNG wire#powerrail
      { S7_Templates := "SrcType := String" } EQ_Contact(in1 := "Expected/Value_All".V, in2 := "Expected/Value_All".Expected_311)
      Move(in := 311, out1 => #Output)
   END_RUNG
   RUNG wire#powerrail
      { S7_Templates := "SrcType := String" } EQ_Contact(in1 := "Expected/Value_All".V, in2 := "Expected/Value_All".Expected_312)
      Move(in := 312, out1 => #Output)
   END_RUNG
   RUNG wire#powerrail
      { S7_Templates := "SrcType := String" } EQ_Contact(in1 := "Expected/Value_All".V, in2 := "Expected/Value_All".Expected_313)
      Move(in := 313, out1 => #Output)
   END_RUNG
   RUNG wire#powerrail
      { S7_Templates := "SrcType := String" } EQ_Contact(in1 := "Expected/Value_All".V, in2 := "Expected/Value_All".Expected_314)
      Move(in := 314, out1 => #Output)
   END_RUNG
   RUNG wire#powerrail
      { S7_Templates := "SrcType := String" } EQ_Contact(in1 := "Expected/Value_All".V, in2 := "Expected/Value_All".Expected_315)
      Move(in := 315, out1 => #Output)
   END_RUNG
   RUNG wire#powerrail
      { S7_Templates := "SrcType := String" } EQ_Contact(in1 := "Expected/Value_All".V, in2 := "Expected/Value_All".Expected_316)
      Move(in := 316, out1 => #Output)
   END_RUNG
   RUNG wire#powerrail
      { S7_Templates := "SrcType := String" } EQ_Contact(in1 := "Expected/Value_All".V, in2 := "Expected/Value_All".Expected_317)
      Move(in := 317, out1 => #Output)
   END_RUNG
   RUNG wire#powerrail
      { S7_Templates := "SrcType := String" } EQ_Contact(in1 := "Expected/Value_All".V, in2 := "Expected/Value_All".Expected_318)
      Move(in := 318, out1 => #Output)
   END_RUNG
   RUNG wire#powerrail
      { S7_Templates := "SrcType := String" } EQ_Contact(in1 := "Expected/Value_All".V, in2 := "Expected/Value_All".Expected_319)
      Move(in := 319, out1 => #Output)
   END_RUNG
   RUNG wire#powerrail
      { S7_Templates := "SrcType := String" } EQ_Contact(in1 := "Expected/Value_All".V, in2 := "Expected/Value_All".Expected_320)
      Move(in := 320, out1 => #Output)
   END_RUNG
   // the same network as SCL:
   IF "Expected/Value_All".V = "Expected/Value_All".Expected_301 THEN #Output := 301; END_IF;
   IF "Expected/Value_All".V = "Expected/Value_All".Expected_302 THEN #Output := 302; END_IF;
   IF "Expected/Value_All".V = "Expected/Value_All".Expected_303 THEN #Output := 303; END_IF;
   IF "Expected/Value_All".V = "Expected/Value_All".Expected_304 THEN #Output := 304; END_IF;
   IF "Expected/Value_All".V = "Expected/Value_All".Expected_305 THEN #Output := 305; END_IF;
   IF "Expected/Value_All".V = "Expected/Value_All".Expected_306 THEN #Output := 306; END_IF;
   IF "Expected/Value_All".V = "Expected/Value_All".Expected_307 THEN #Output := 307; END_IF;
   IF "Expected/Value_All".V = "Expected/Value_All".Expected_308 THEN #Output := 308; END_IF;
   IF "Expected/Value_All".V = "Expected/Value_All".Expected_309 THEN #Output := 309; END_IF;
   IF "Expected/Value_All".V = "Expected/Value_All".Expected_310 THEN #Output := 310; END_IF;
   IF "Expected/Value_All".V = "Expected/Value_All".Expected_311 THEN #Output := 311; END_IF;
   IF "Expected/Value_All".V = "Expected/Value_All".Expected_312 THEN #Output := 312; END_IF;
   IF "Expected/Value_All".V = "Expected/Value_All".Expected_313 THEN #Output := 313; END_IF;
   IF "Expected/Value_All".V = "Expected/Value_All".Expected_314 THEN #Output := 314; END_IF;
   IF "Expected/Value_All".V = "Expected/Value_All".Expected_315 THEN #Output := 315; END_IF;
   IF "Expected/Value_All".V = "Expected/Value_All".Expected_316 THEN #Output := 316; END_IF;
   IF "Expected/Value_All".V = "Expected/Value_All".Expected_317 THEN #Output := 317; END_IF;
   IF "Expected/Value_All".V = "Expected/Value_All".Expected_318 THEN #Output := 318; END_IF;
   IF "Expected/Value_All".V = "Expected/Value_All".Expected_319 THEN #Output := 319; END_IF;
   IF "Expected/Value_All".V = "Expected/Value_All".Expected_320 THEN #Output := 320; END_IF;
END_REGION

REGION Network 17
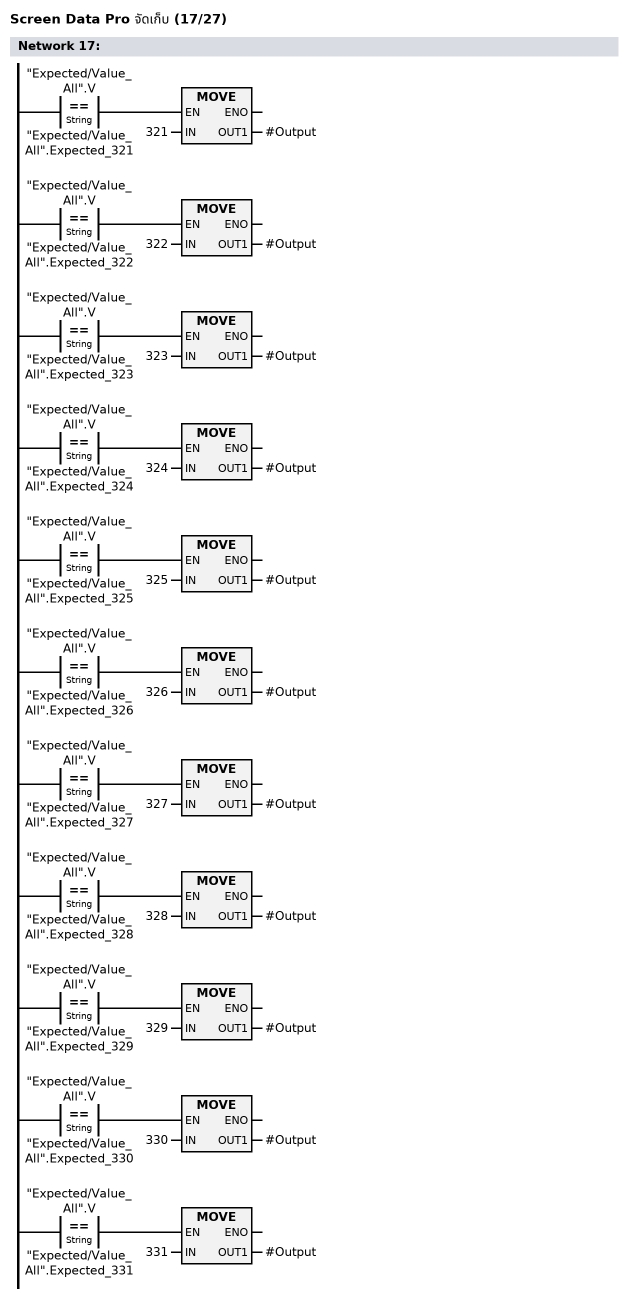
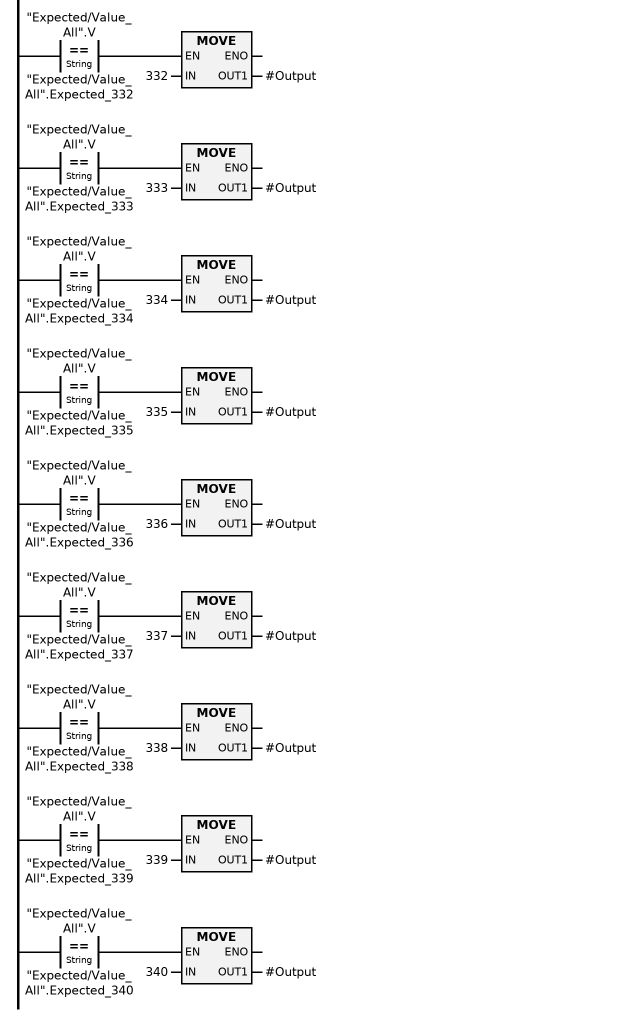
   RUNG wire#powerrail
      { S7_Templates := "SrcType := String" } EQ_Contact(in1 := "Expected/Value_All".V, in2 := "Expected/Value_All".Expected_321)
      Move(in := 321, out1 => #Output)
   END_RUNG
   RUNG wire#powerrail
      { S7_Templates := "SrcType := String" } EQ_Contact(in1 := "Expected/Value_All".V, in2 := "Expected/Value_All".Expected_322)
      Move(in := 322, out1 => #Output)
   END_RUNG
   RUNG wire#powerrail
      { S7_Templates := "SrcType := String" } EQ_Contact(in1 := "Expected/Value_All".V, in2 := "Expected/Value_All".Expected_323)
      Move(in := 323, out1 => #Output)
   END_RUNG
   RUNG wire#powerrail
      { S7_Templates := "SrcType := String" } EQ_Contact(in1 := "Expected/Value_All".V, in2 := "Expected/Value_All".Expected_324)
      Move(in := 324, out1 => #Output)
   END_RUNG
   RUNG wire#powerrail
      { S7_Templates := "SrcType := String" } EQ_Contact(in1 := "Expected/Value_All".V, in2 := "Expected/Value_All".Expected_325)
      Move(in := 325, out1 => #Output)
   END_RUNG
   RUNG wire#powerrail
      { S7_Templates := "SrcType := String" } EQ_Contact(in1 := "Expected/Value_All".V, in2 := "Expected/Value_All".Expected_326)
      Move(in := 326, out1 => #Output)
   END_RUNG
   RUNG wire#powerrail
      { S7_Templates := "SrcType := String" } EQ_Contact(in1 := "Expected/Value_All".V, in2 := "Expected/Value_All".Expected_327)
      Move(in := 327, out1 => #Output)
   END_RUNG
   RUNG wire#powerrail
      { S7_Templates := "SrcType := String" } EQ_Contact(in1 := "Expected/Value_All".V, in2 := "Expected/Value_All".Expected_328)
      Move(in := 328, out1 => #Output)
   END_RUNG
   RUNG wire#powerrail
      { S7_Templates := "SrcType := String" } EQ_Contact(in1 := "Expected/Value_All".V, in2 := "Expected/Value_All".Expected_329)
      Move(in := 329, out1 => #Output)
   END_RUNG
   RUNG wire#powerrail
      { S7_Templates := "SrcType := String" } EQ_Contact(in1 := "Expected/Value_All".V, in2 := "Expected/Value_All".Expected_330)
      Move(in := 330, out1 => #Output)
   END_RUNG
   RUNG wire#powerrail
      { S7_Templates := "SrcType := String" } EQ_Contact(in1 := "Expected/Value_All".V, in2 := "Expected/Value_All".Expected_331)
      Move(in := 331, out1 => #Output)
   END_RUNG
   RUNG wire#powerrail
      { S7_Templates := "SrcType := String" } EQ_Contact(in1 := "Expected/Value_All".V, in2 := "Expected/Value_All".Expected_332)
      Move(in := 332, out1 => #Output)
   END_RUNG
   RUNG wire#powerrail
      { S7_Templates := "SrcType := String" } EQ_Contact(in1 := "Expected/Value_All".V, in2 := "Expected/Value_All".Expected_333)
      Move(in := 333, out1 => #Output)
   END_RUNG
   RUNG wire#powerrail
      { S7_Templates := "SrcType := String" } EQ_Contact(in1 := "Expected/Value_All".V, in2 := "Expected/Value_All".Expected_334)
      Move(in := 334, out1 => #Output)
   END_RUNG
   RUNG wire#powerrail
      { S7_Templates := "SrcType := String" } EQ_Contact(in1 := "Expected/Value_All".V, in2 := "Expected/Value_All".Expected_335)
      Move(in := 335, out1 => #Output)
   END_RUNG
   RUNG wire#powerrail
      { S7_Templates := "SrcType := String" } EQ_Contact(in1 := "Expected/Value_All".V, in2 := "Expected/Value_All".Expected_336)
      Move(in := 336, out1 => #Output)
   END_RUNG
   RUNG wire#powerrail
      { S7_Templates := "SrcType := String" } EQ_Contact(in1 := "Expected/Value_All".V, in2 := "Expected/Value_All".Expected_337)
      Move(in := 337, out1 => #Output)
   END_RUNG
   RUNG wire#powerrail
      { S7_Templates := "SrcType := String" } EQ_Contact(in1 := "Expected/Value_All".V, in2 := "Expected/Value_All".Expected_338)
      Move(in := 338, out1 => #Output)
   END_RUNG
   RUNG wire#powerrail
      { S7_Templates := "SrcType := String" } EQ_Contact(in1 := "Expected/Value_All".V, in2 := "Expected/Value_All".Expected_339)
      Move(in := 339, out1 => #Output)
   END_RUNG
   RUNG wire#powerrail
      { S7_Templates := "SrcType := String" } EQ_Contact(in1 := "Expected/Value_All".V, in2 := "Expected/Value_All".Expected_340)
      Move(in := 340, out1 => #Output)
   END_RUNG
   // the same network as SCL:
   IF "Expected/Value_All".V = "Expected/Value_All".Expected_321 THEN #Output := 321; END_IF;
   IF "Expected/Value_All".V = "Expected/Value_All".Expected_322 THEN #Output := 322; END_IF;
   IF "Expected/Value_All".V = "Expected/Value_All".Expected_323 THEN #Output := 323; END_IF;
   IF "Expected/Value_All".V = "Expected/Value_All".Expected_324 THEN #Output := 324; END_IF;
   IF "Expected/Value_All".V = "Expected/Value_All".Expected_325 THEN #Output := 325; END_IF;
   IF "Expected/Value_All".V = "Expected/Value_All".Expected_326 THEN #Output := 326; END_IF;
   IF "Expected/Value_All".V = "Expected/Value_All".Expected_327 THEN #Output := 327; END_IF;
   IF "Expected/Value_All".V = "Expected/Value_All".Expected_328 THEN #Output := 328; END_IF;
   IF "Expected/Value_All".V = "Expected/Value_All".Expected_329 THEN #Output := 329; END_IF;
   IF "Expected/Value_All".V = "Expected/Value_All".Expected_330 THEN #Output := 330; END_IF;
   IF "Expected/Value_All".V = "Expected/Value_All".Expected_331 THEN #Output := 331; END_IF;
   IF "Expected/Value_All".V = "Expected/Value_All".Expected_332 THEN #Output := 332; END_IF;
   IF "Expected/Value_All".V = "Expected/Value_All".Expected_333 THEN #Output := 333; END_IF;
   IF "Expected/Value_All".V = "Expected/Value_All".Expected_334 THEN #Output := 334; END_IF;
   IF "Expected/Value_All".V = "Expected/Value_All".Expected_335 THEN #Output := 335; END_IF;
   IF "Expected/Value_All".V = "Expected/Value_All".Expected_336 THEN #Output := 336; END_IF;
   IF "Expected/Value_All".V = "Expected/Value_All".Expected_337 THEN #Output := 337; END_IF;
   IF "Expected/Value_All".V = "Expected/Value_All".Expected_338 THEN #Output := 338; END_IF;
   IF "Expected/Value_All".V = "Expected/Value_All".Expected_339 THEN #Output := 339; END_IF;
   IF "Expected/Value_All".V = "Expected/Value_All".Expected_340 THEN #Output := 340; END_IF;
END_REGION

REGION Network 18
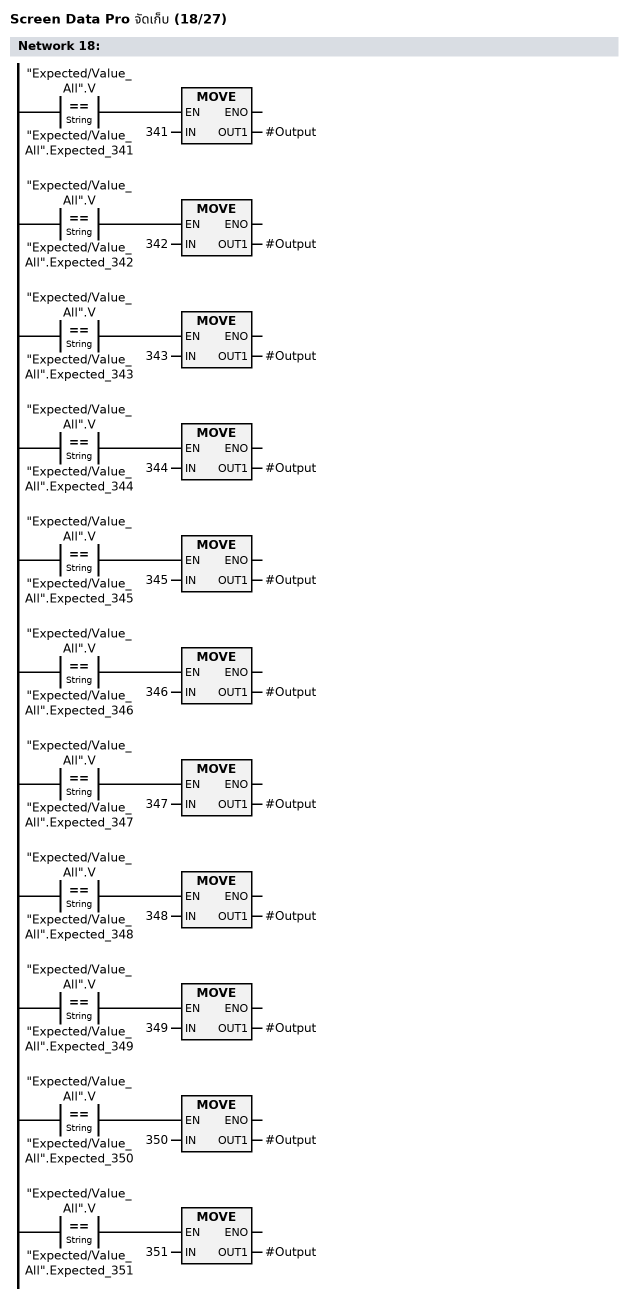
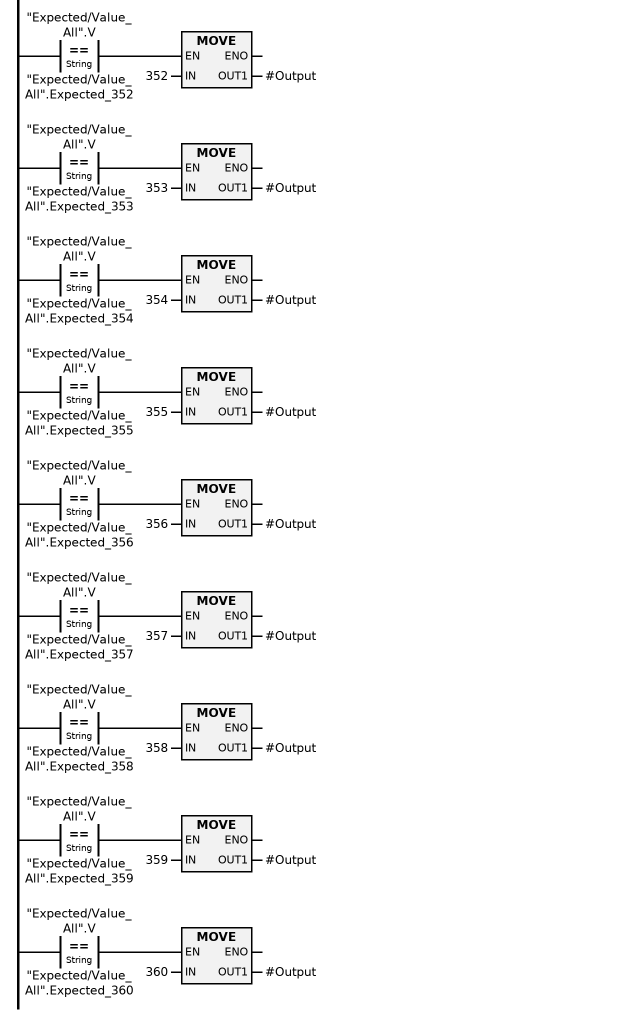
   RUNG wire#powerrail
      { S7_Templates := "SrcType := String" } EQ_Contact(in1 := "Expected/Value_All".V, in2 := "Expected/Value_All".Expected_341)
      Move(in := 341, out1 => #Output)
   END_RUNG
   RUNG wire#powerrail
      { S7_Templates := "SrcType := String" } EQ_Contact(in1 := "Expected/Value_All".V, in2 := "Expected/Value_All".Expected_342)
      Move(in := 342, out1 => #Output)
   END_RUNG
   RUNG wire#powerrail
      { S7_Templates := "SrcType := String" } EQ_Contact(in1 := "Expected/Value_All".V, in2 := "Expected/Value_All".Expected_343)
      Move(in := 343, out1 => #Output)
   END_RUNG
   RUNG wire#powerrail
      { S7_Templates := "SrcType := String" } EQ_Contact(in1 := "Expected/Value_All".V, in2 := "Expected/Value_All".Expected_344)
      Move(in := 344, out1 => #Output)
   END_RUNG
   RUNG wire#powerrail
      { S7_Templates := "SrcType := String" } EQ_Contact(in1 := "Expected/Value_All".V, in2 := "Expected/Value_All".Expected_345)
      Move(in := 345, out1 => #Output)
   END_RUNG
   RUNG wire#powerrail
      { S7_Templates := "SrcType := String" } EQ_Contact(in1 := "Expected/Value_All".V, in2 := "Expected/Value_All".Expected_346)
      Move(in := 346, out1 => #Output)
   END_RUNG
   RUNG wire#powerrail
      { S7_Templates := "SrcType := String" } EQ_Contact(in1 := "Expected/Value_All".V, in2 := "Expected/Value_All".Expected_347)
      Move(in := 347, out1 => #Output)
   END_RUNG
   RUNG wire#powerrail
      { S7_Templates := "SrcType := String" } EQ_Contact(in1 := "Expected/Value_All".V, in2 := "Expected/Value_All".Expected_348)
      Move(in := 348, out1 => #Output)
   END_RUNG
   RUNG wire#powerrail
      { S7_Templates := "SrcType := String" } EQ_Contact(in1 := "Expected/Value_All".V, in2 := "Expected/Value_All".Expected_349)
      Move(in := 349, out1 => #Output)
   END_RUNG
   RUNG wire#powerrail
      { S7_Templates := "SrcType := String" } EQ_Contact(in1 := "Expected/Value_All".V, in2 := "Expected/Value_All".Expected_350)
      Move(in := 350, out1 => #Output)
   END_RUNG
   RUNG wire#powerrail
      { S7_Templates := "SrcType := String" } EQ_Contact(in1 := "Expected/Value_All".V, in2 := "Expected/Value_All".Expected_351)
      Move(in := 351, out1 => #Output)
   END_RUNG
   RUNG wire#powerrail
      { S7_Templates := "SrcType := String" } EQ_Contact(in1 := "Expected/Value_All".V, in2 := "Expected/Value_All".Expected_352)
      Move(in := 352, out1 => #Output)
   END_RUNG
   RUNG wire#powerrail
      { S7_Templates := "SrcType := String" } EQ_Contact(in1 := "Expected/Value_All".V, in2 := "Expected/Value_All".Expected_353)
      Move(in := 353, out1 => #Output)
   END_RUNG
   RUNG wire#powerrail
      { S7_Templates := "SrcType := String" } EQ_Contact(in1 := "Expected/Value_All".V, in2 := "Expected/Value_All".Expected_354)
      Move(in := 354, out1 => #Output)
   END_RUNG
   RUNG wire#powerrail
      { S7_Templates := "SrcType := String" } EQ_Contact(in1 := "Expected/Value_All".V, in2 := "Expected/Value_All".Expected_355)
      Move(in := 355, out1 => #Output)
   END_RUNG
   RUNG wire#powerrail
      { S7_Templates := "SrcType := String" } EQ_Contact(in1 := "Expected/Value_All".V, in2 := "Expected/Value_All".Expected_356)
      Move(in := 356, out1 => #Output)
   END_RUNG
   RUNG wire#powerrail
      { S7_Templates := "SrcType := String" } EQ_Contact(in1 := "Expected/Value_All".V, in2 := "Expected/Value_All".Expected_357)
      Move(in := 357, out1 => #Output)
   END_RUNG
   RUNG wire#powerrail
      { S7_Templates := "SrcType := String" } EQ_Contact(in1 := "Expected/Value_All".V, in2 := "Expected/Value_All".Expected_358)
      Move(in := 358, out1 => #Output)
   END_RUNG
   RUNG wire#powerrail
      { S7_Templates := "SrcType := String" } EQ_Contact(in1 := "Expected/Value_All".V, in2 := "Expected/Value_All".Expected_359)
      Move(in := 359, out1 => #Output)
   END_RUNG
   RUNG wire#powerrail
      { S7_Templates := "SrcType := String" } EQ_Contact(in1 := "Expected/Value_All".V, in2 := "Expected/Value_All".Expected_360)
      Move(in := 360, out1 => #Output)
   END_RUNG
   // the same network as SCL:
   IF "Expected/Value_All".V = "Expected/Value_All".Expected_341 THEN #Output := 341; END_IF;
   IF "Expected/Value_All".V = "Expected/Value_All".Expected_342 THEN #Output := 342; END_IF;
   IF "Expected/Value_All".V = "Expected/Value_All".Expected_343 THEN #Output := 343; END_IF;
   IF "Expected/Value_All".V = "Expected/Value_All".Expected_344 THEN #Output := 344; END_IF;
   IF "Expected/Value_All".V = "Expected/Value_All".Expected_345 THEN #Output := 345; END_IF;
   IF "Expected/Value_All".V = "Expected/Value_All".Expected_346 THEN #Output := 346; END_IF;
   IF "Expected/Value_All".V = "Expected/Value_All".Expected_347 THEN #Output := 347; END_IF;
   IF "Expected/Value_All".V = "Expected/Value_All".Expected_348 THEN #Output := 348; END_IF;
   IF "Expected/Value_All".V = "Expected/Value_All".Expected_349 THEN #Output := 349; END_IF;
   IF "Expected/Value_All".V = "Expected/Value_All".Expected_350 THEN #Output := 350; END_IF;
   IF "Expected/Value_All".V = "Expected/Value_All".Expected_351 THEN #Output := 351; END_IF;
   IF "Expected/Value_All".V = "Expected/Value_All".Expected_352 THEN #Output := 352; END_IF;
   IF "Expected/Value_All".V = "Expected/Value_All".Expected_353 THEN #Output := 353; END_IF;
   IF "Expected/Value_All".V = "Expected/Value_All".Expected_354 THEN #Output := 354; END_IF;
   IF "Expected/Value_All".V = "Expected/Value_All".Expected_355 THEN #Output := 355; END_IF;
   IF "Expected/Value_All".V = "Expected/Value_All".Expected_356 THEN #Output := 356; END_IF;
   IF "Expected/Value_All".V = "Expected/Value_All".Expected_357 THEN #Output := 357; END_IF;
   IF "Expected/Value_All".V = "Expected/Value_All".Expected_358 THEN #Output := 358; END_IF;
   IF "Expected/Value_All".V = "Expected/Value_All".Expected_359 THEN #Output := 359; END_IF;
   IF "Expected/Value_All".V = "Expected/Value_All".Expected_360 THEN #Output := 360; END_IF;
END_REGION

REGION Network 19
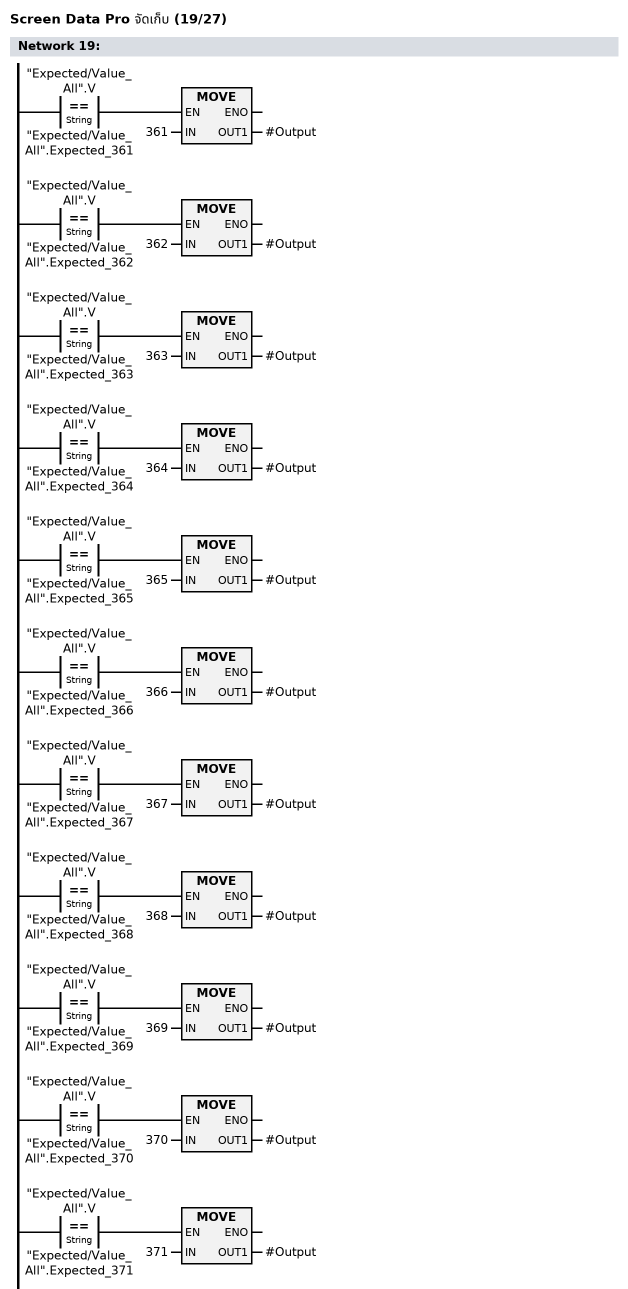
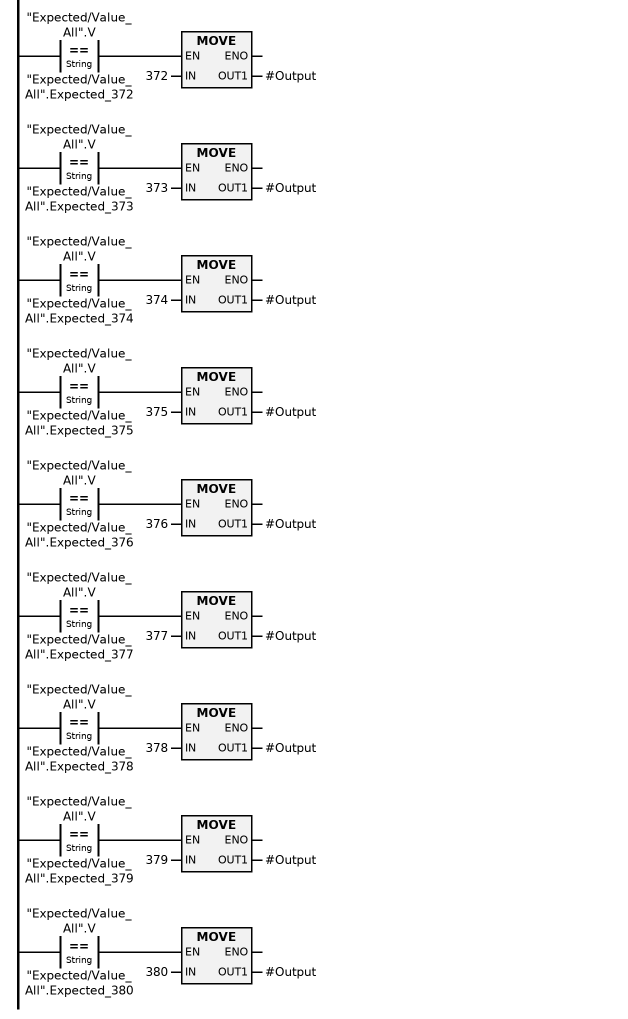
   RUNG wire#powerrail
      { S7_Templates := "SrcType := String" } EQ_Contact(in1 := "Expected/Value_All".V, in2 := "Expected/Value_All".Expected_361)
      Move(in := 361, out1 => #Output)
   END_RUNG
   RUNG wire#powerrail
      { S7_Templates := "SrcType := String" } EQ_Contact(in1 := "Expected/Value_All".V, in2 := "Expected/Value_All".Expected_362)
      Move(in := 362, out1 => #Output)
   END_RUNG
   RUNG wire#powerrail
      { S7_Templates := "SrcType := String" } EQ_Contact(in1 := "Expected/Value_All".V, in2 := "Expected/Value_All".Expected_363)
      Move(in := 363, out1 => #Output)
   END_RUNG
   RUNG wire#powerrail
      { S7_Templates := "SrcType := String" } EQ_Contact(in1 := "Expected/Value_All".V, in2 := "Expected/Value_All".Expected_364)
      Move(in := 364, out1 => #Output)
   END_RUNG
   RUNG wire#powerrail
      { S7_Templates := "SrcType := String" } EQ_Contact(in1 := "Expected/Value_All".V, in2 := "Expected/Value_All".Expected_365)
      Move(in := 365, out1 => #Output)
   END_RUNG
   RUNG wire#powerrail
      { S7_Templates := "SrcType := String" } EQ_Contact(in1 := "Expected/Value_All".V, in2 := "Expected/Value_All".Expected_366)
      Move(in := 366, out1 => #Output)
   END_RUNG
   RUNG wire#powerrail
      { S7_Templates := "SrcType := String" } EQ_Contact(in1 := "Expected/Value_All".V, in2 := "Expected/Value_All".Expected_367)
      Move(in := 367, out1 => #Output)
   END_RUNG
   RUNG wire#powerrail
      { S7_Templates := "SrcType := String" } EQ_Contact(in1 := "Expected/Value_All".V, in2 := "Expected/Value_All".Expected_368)
      Move(in := 368, out1 => #Output)
   END_RUNG
   RUNG wire#powerrail
      { S7_Templates := "SrcType := String" } EQ_Contact(in1 := "Expected/Value_All".V, in2 := "Expected/Value_All".Expected_369)
      Move(in := 369, out1 => #Output)
   END_RUNG
   RUNG wire#powerrail
      { S7_Templates := "SrcType := String" } EQ_Contact(in1 := "Expected/Value_All".V, in2 := "Expected/Value_All".Expected_370)
      Move(in := 370, out1 => #Output)
   END_RUNG
   RUNG wire#powerrail
      { S7_Templates := "SrcType := String" } EQ_Contact(in1 := "Expected/Value_All".V, in2 := "Expected/Value_All".Expected_371)
      Move(in := 371, out1 => #Output)
   END_RUNG
   RUNG wire#powerrail
      { S7_Templates := "SrcType := String" } EQ_Contact(in1 := "Expected/Value_All".V, in2 := "Expected/Value_All".Expected_372)
      Move(in := 372, out1 => #Output)
   END_RUNG
   RUNG wire#powerrail
      { S7_Templates := "SrcType := String" } EQ_Contact(in1 := "Expected/Value_All".V, in2 := "Expected/Value_All".Expected_373)
      Move(in := 373, out1 => #Output)
   END_RUNG
   RUNG wire#powerrail
      { S7_Templates := "SrcType := String" } EQ_Contact(in1 := "Expected/Value_All".V, in2 := "Expected/Value_All".Expected_374)
      Move(in := 374, out1 => #Output)
   END_RUNG
   RUNG wire#powerrail
      { S7_Templates := "SrcType := String" } EQ_Contact(in1 := "Expected/Value_All".V, in2 := "Expected/Value_All".Expected_375)
      Move(in := 375, out1 => #Output)
   END_RUNG
   RUNG wire#powerrail
      { S7_Templates := "SrcType := String" } EQ_Contact(in1 := "Expected/Value_All".V, in2 := "Expected/Value_All".Expected_376)
      Move(in := 376, out1 => #Output)
   END_RUNG
   RUNG wire#powerrail
      { S7_Templates := "SrcType := String" } EQ_Contact(in1 := "Expected/Value_All".V, in2 := "Expected/Value_All".Expected_377)
      Move(in := 377, out1 => #Output)
   END_RUNG
   RUNG wire#powerrail
      { S7_Templates := "SrcType := String" } EQ_Contact(in1 := "Expected/Value_All".V, in2 := "Expected/Value_All".Expected_378)
      Move(in := 378, out1 => #Output)
   END_RUNG
   RUNG wire#powerrail
      { S7_Templates := "SrcType := String" } EQ_Contact(in1 := "Expected/Value_All".V, in2 := "Expected/Value_All".Expected_379)
      Move(in := 379, out1 => #Output)
   END_RUNG
   RUNG wire#powerrail
      { S7_Templates := "SrcType := String" } EQ_Contact(in1 := "Expected/Value_All".V, in2 := "Expected/Value_All".Expected_380)
      Move(in := 380, out1 => #Output)
   END_RUNG
   // the same network as SCL:
   IF "Expected/Value_All".V = "Expected/Value_All".Expected_361 THEN #Output := 361; END_IF;
   IF "Expected/Value_All".V = "Expected/Value_All".Expected_362 THEN #Output := 362; END_IF;
   IF "Expected/Value_All".V = "Expected/Value_All".Expected_363 THEN #Output := 363; END_IF;
   IF "Expected/Value_All".V = "Expected/Value_All".Expected_364 THEN #Output := 364; END_IF;
   IF "Expected/Value_All".V = "Expected/Value_All".Expected_365 THEN #Output := 365; END_IF;
   IF "Expected/Value_All".V = "Expected/Value_All".Expected_366 THEN #Output := 366; END_IF;
   IF "Expected/Value_All".V = "Expected/Value_All".Expected_367 THEN #Output := 367; END_IF;
   IF "Expected/Value_All".V = "Expected/Value_All".Expected_368 THEN #Output := 368; END_IF;
   IF "Expected/Value_All".V = "Expected/Value_All".Expected_369 THEN #Output := 369; END_IF;
   IF "Expected/Value_All".V = "Expected/Value_All".Expected_370 THEN #Output := 370; END_IF;
   IF "Expected/Value_All".V = "Expected/Value_All".Expected_371 THEN #Output := 371; END_IF;
   IF "Expected/Value_All".V = "Expected/Value_All".Expected_372 THEN #Output := 372; END_IF;
   IF "Expected/Value_All".V = "Expected/Value_All".Expected_373 THEN #Output := 373; END_IF;
   IF "Expected/Value_All".V = "Expected/Value_All".Expected_374 THEN #Output := 374; END_IF;
   IF "Expected/Value_All".V = "Expected/Value_All".Expected_375 THEN #Output := 375; END_IF;
   IF "Expected/Value_All".V = "Expected/Value_All".Expected_376 THEN #Output := 376; END_IF;
   IF "Expected/Value_All".V = "Expected/Value_All".Expected_377 THEN #Output := 377; END_IF;
   IF "Expected/Value_All".V = "Expected/Value_All".Expected_378 THEN #Output := 378; END_IF;
   IF "Expected/Value_All".V = "Expected/Value_All".Expected_379 THEN #Output := 379; END_IF;
   IF "Expected/Value_All".V = "Expected/Value_All".Expected_380 THEN #Output := 380; END_IF;
END_REGION

REGION Network 20
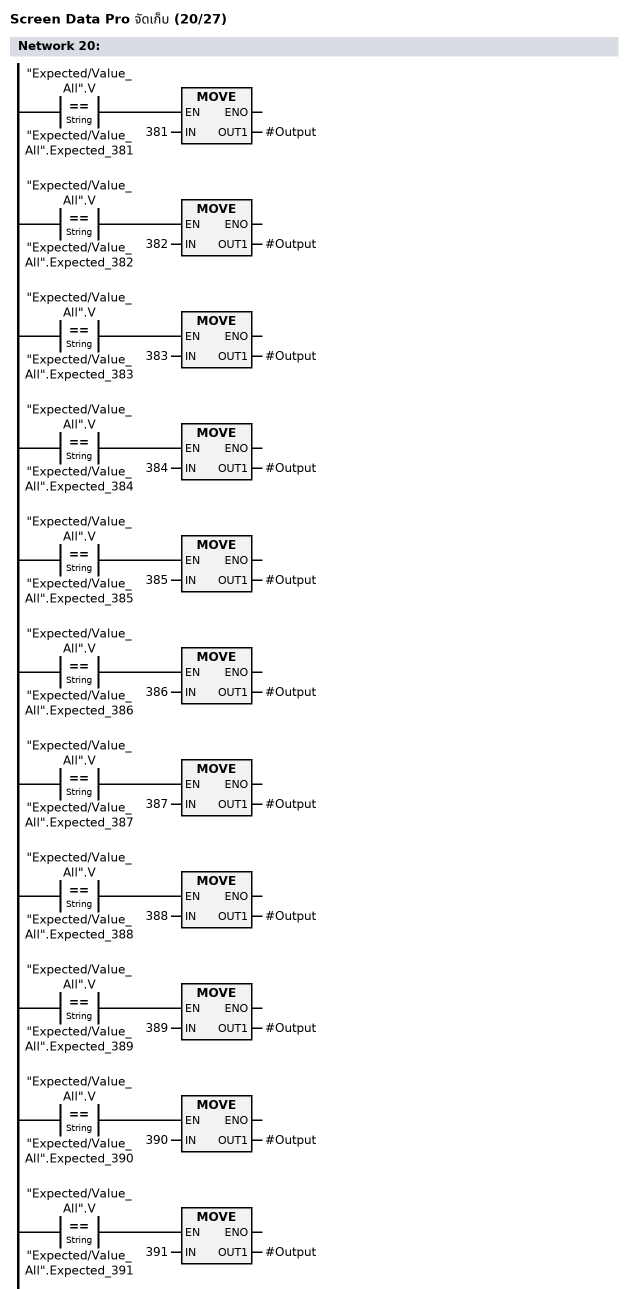
